(* IEC 61131-3 sources: 2026_Projet_YGO_ExcavatriceDragage/CODE/L_SIMULATION, 12 files *)

(* ---- FB_Sim_Encoder.st ---- *)
(* ═══════════════════════════════════════════════════════════════
   🧪 FB_Sim_Encoder — Simulation physique d'un codeur absolu de treuil
   ───────────────────────────────────────────────────────────────
   📄 Doc métier : DOC/AF/AF_Partie-13_Fonction_Simulation_v2.5.md
   📄 Spec composant : DOC/AF/AF_Partie-13_Fonction_Simulation/FB_Sim_Encoder_v1.1.md
   🧩 Brique réduite (Partie3 §1bis, "briques E/S & diagnostics") : pas de contrat
      Enable/Reset/Error complet, pas de StartStop/SafeStop — outil de banc, pas
      du métier machine.
   🎯 Rôle : fait "compter" un codeur absolu comme si le treuil tournait
      réellement, à partir des relais de sens commandés et du palier de vitesse courant.
   📥 Enable      : simulation active (SimulationModeActive AND NOT BusEncoderMxIsReal)
   📥 RelayFwd/RelayRev : sens commandé (contacteurs de sens du treuil)
   📥 StepNumber  : palier vitesse courant (1..5) — ex. instWinchM1.StepNumber
      Vitesse = interpolation linéaire : palier 1 → MinSpeedMps (1 m/s), palier 5 → MaxSpeedMps (2 m/s).
   📥 PresetCmd   : TRUE le cycle où un preset (homing) doit être appliqué (PresettTrigCmd = 2)
   📥 PresetValue : valeur brute à charger lors du preset
   📥 SpeedScaleFactor : facteur fin de confort (réglable à chaud, sans recompiler). Défaut 1.0 = vitesse
      réelle telle que définie par MinSpeedMps/MaxSpeedMps/PointsPerRev/CableM_PerRev/CycleTimeS.
   📤 RawPosOut   : position brute simulée (UDINT), à aiguiller à la place de la valeur
      EtherCAT réelle quand le device n'est pas Operational (voir PRG_02_Encoders.st)
   🔒 Comptage brut : entier SIGNÉ 32 bits (le conteneur UDINT n'est qu'un support d'échange,
      relu en DINT par toute la chaîne aval). Il franchit 0 sans jamais s'y figer ; la seule
      borne est la plage de représentation, signalée par CountSaturated — jamais muette.
   📤 CountSaturated : comptage en butée de plage du modèle (saturation signalée, vitesse purgée)
   `RawPos` en `VAR_IN_OUT`, référencé depuis `GVL_PERSISTENT`
      (même pattern que `Calib` dans `FB_Encoder_Homing`) — `PERSISTENT` n'est valide que sur du
      `VAR_GLOBAL` en CODESYS, pas sur une variable locale de FB. Un vrai codeur absolu physique
      conserve son comptage brut même à travers un reset FROID (indépendant de l'automate).
   ═══════════════════════════════════════════════════════════════ *)

// === DECLARATION (à coller dans la partie déclaration du POU FB_Sim_Encoder) ===

FUNCTION_BLOCK PUBLIC FB_Sim_Encoder
VAR_INPUT
    Enable           : BOOL;   (* --> [CMD] Active la simulation *)
    RelayFwd         : BOOL;   (* --> [HW] Sens commandé avant *)
    RelayRev         : BOOL;   (* --> [HW] Sens commandé arrière *)
    StepNumber       : INT;    (* --> [CMD] Palier vitesse courant (1..5, 0 = arrêt) *)
    PresetCmd        : BOOL;   (* --> [CMD] Applique un preset (homing) *)
    PresetValue      : UDINT;   (* --> [CFG] Valeur brute à charger au preset *)
    SpeedScaleFactor : REAL := 1.0;   (* --> [CFG] Facteur fin de confort (défaut 1.0) *)
    CoastDistanceM   : REAL := 0.0;   (* --> [CFG] Distance de roulis inertiel apres coupure des relais (m). 0 = arret net (defaut). >0 = le treuil continue a vitesse palier 1 dans le dernier sens sur CoastDistanceM metres -> modelise l'anticipation d'arret mecanique (ex. benne). *)
    PresetLatencyCycles : INT := 3;   (* --> [CFG] Nb cycles automate avant application du preset (referencement non instantane) *)
    TestOffsetCmd    : BOOL;          (* --> [TST] Front montant = applique TestOffsetPts (test banc) *)
    TestOffsetPts    : DINT := 0;     (* --> [TST] Décalage signé à appliquer (points bruts) *)
    // 📐 Paramètres physiques du treuil (mêmes valeurs que FB_Encoder_Scale) + vitesse réelle.
    // Vitesse simulée = interpolation linéaire du palier : palier 1 → MinSpeedMps, palier 5 → MaxSpeedMps.
    MinSpeedMps      : REAL := 1.0;    (* --> [CFG] Vitesse palier 1 (m/s) *)
    MaxSpeedMps      : REAL := 2.0;    (* --> [CFG] Vitesse palier 5 (m/s) *)
    PointsPerRev     : UDINT := 8192;  (* --> [CFG] Résolution codeur (pts/tour) *)
    CableM_PerRev    : REAL := 2.0;    (* --> [CFG] Développement câble (m/tour) *)
    CycleTimeS       : REAL := 0.010;  (* --> [CFG] Période tâche PLC (s) — MainTask 10 ms *)
    SpeedReportTauS  : REAL := 0.0;    (* --> [CFG][SYNTHETIQUE] Constante de temps 1er ordre du retour vitesse
        (RawSpdOut), s. 0.0 = saut instantane. >0 = RawSpdOut suit un 1er ordre vers la vitesse reelle du modele
        au lieu de sauter en escalier a la coupure des relais ; RawPosOut (position) n'est pas affecte. Valeur
        non calibree treuil M1/M2, plage indicative issue de la dynamique variateur M3 identifiee sur trace. *)
    // 🆕 Dynamique de glissement inertiel fidele (T421 cale sur trace reelle Suivi_86)
    CoastDecelUp_Mps2   : REAL := 1.20;  (* --> [CFG] Deceleration en montee (m/s²) : v0²/(2*0.543m) = 1.20 *)
    CoastDecelDown_Mps2 : REAL := 0.93;  (* --> [CFG] Deceleration en descente (m/s²) : v0²/(2*1.205m) = 0.93 *)
    MechanicStopEngaged : BOOL := FALSE; (* --> [HW] Butee mecanique engagee (coupe net le glissement) *)
END_VAR
VAR_OUTPUT
    RawPosOut   : UDINT;   (* <-- [DIAG] Position brute simulée *)
    RawSpdOut   : DINT;    (* <-- [DIAG] Vitesse brute simulée (0x6031:01 en 0.1 RPM) *)
    CountSaturated : BOOL; (* <-- [DIAG] Comptage en butée de plage du modèle (saturation signalée) *)
    CoastActive    : BOOL; (* <-- [DIAG] Indicateur de glissement inertiel en cours (T421) *)
END_VAR
VAR_IN_OUT
    RawPos      : UDINT;   (* <-> [BUS] Référence _SimEncoderRawPosM1/M2 (survit au reset froid) *)
END_VAR
VAR
    Increment        : UDINT;            (* . [LOC] Points ajoutés par cycle *)
    EffStep          : INT;              (* . [LOC] Pas borné (>= 1) *)
    SpeedMps         : REAL;             (* . [LOC] Vitesse simulée (m/s) *)
    TestOffsetEdge   : R_TRIG;           (* . [LOC] Front TestOffsetCmd *)
    PresetEdge       : R_TRIG;           (* . [LOC] Front montant PresetCmd *)
    PresetPending    : BOOL;             (* . [LOC] Preset en attente d'application (latence) *)
    PresetCount      : INT;              (* . [LOC] Compteur cycles de latence restants *)
    IncrStep1        : UDINT;            (* . [LOC] Increment par cycle a vitesse palier 1 (pour le roulis) *)
    MovingDir        : INT;              (* . [LOC] Dernier sens actif : +1 avant, -1 arriere, 0 arret *)
    CoastPtsLeft     : REAL;             (* . [LOC] Roulis inertiel restant (points bruts) *)
    TargetSpeedMps   : REAL;             (* . [LOC] Vitesse instantanee signee du modele position, avant filtrage retour *)
    ReportedSpeedMps : REAL;             (* . [LOC] Vitesse rapportee filtree 1er ordre, publiee dans RawSpdOut *)
    CoastSpeedMps    : REAL;             (* . [LOC] Vitesse instantanee signee pendant le glissement inertiel (T421) *)
END_VAR
VAR CONSTANT
    // 🛑 Plage de comptage du modèle : le compteur brut est un entier SIGNÉ 32 bits (le conteneur
    // UDINT n'est qu'un support d'échange, relu en DINT par toute la chaîne aval). La garde reste
    // volontairement à la moitié de la plage signée (2^30 pts = 262 144 m de câble) : inatteignable
    // en essai, elle interdit tout rebouclage silencieux si le modèle consommait toute sa plage.
    CST_CountTravelLimitPts : DINT := 1073741824; // 2^30 pts — demi-plage signée
END_VAR

// === IMPLEMENTATION (à coller dans le corps ST du POU FB_Sim_Encoder) ===

{region "§1 Gate"}
IF NOT Enable THEN
    RawPosOut := RawPos;
    // Comptage non evalue hors simulation : la saturation ne doit pas rester figee a TRUE.
    CountSaturated := FALSE;
    RETURN;
END_IF;
{endregion}

{region "§2 Injection test"}
// Injection test banc : VRAI saut de position (comme un glissement réel),
// pour tester Concept 1 / Méca E ET le rattrapage joystick (voir GVL_Simulation bandeau).
TestOffsetEdge(CLK := TestOffsetCmd);
IF TestOffsetEdge.Q THEN
    RawPos := DINT_TO_UDINT(UDINT_TO_DINT(RawPos) + TestOffsetPts);
END_IF;
{endregion}

{region "§3 Comptage"}
// 🎚️ Vitesse simulée = interpolation linéaire du palier (palier 1 → MinSpeedMps, palier 5 → MaxSpeedMps),
// pas par pas de (Max−Min)/4. Palier 0 (arrêt) ramène au palier 1 mais aucun mouvement n'est
// appliqué tant que RelayFwd/RelayRev = FALSE (section plus bas).
EffStep  := MAX(StepNumber, 1);
SpeedMps := MinSpeedMps + (INT_TO_REAL(EffStep) - 1.0) * ((MaxSpeedMps - MinSpeedMps) / 4.0);
// Points par cycle = vitesse (m/s) × points par mètre × période tâche (s) × facteur confort.
Increment := REAL_TO_UDINT(SpeedMps * (UDINT_TO_REAL(PointsPerRev) / CableM_PerRev) * CycleTimeS * SpeedScaleFactor);
// Increment "lent" (palier 1) : vitesse du roulis inertiel apres coupure des relais.
IncrStep1 := REAL_TO_UDINT(MinSpeedMps * (UDINT_TO_REAL(PointsPerRev) / CableM_PerRev) * CycleTimeS * SpeedScaleFactor);

// Front du preset : lance la latence de referencement (le codeur réel n'est pas
// instantane — il met PresetLatencyCycles cycles a se re-referencer apres le front).
PresetEdge(CLK := PresetCmd);
IF PresetEdge.Q THEN
    PresetPending := TRUE;
    PresetCount := PresetLatencyCycles;
END_IF;

// 📐 Le comptage brut est un entier SIGNÉ 32 bits : le conteneur UDINT n'est qu'un support
// d'échange (toute la chaîne aval le relit via UDINT_TO_DINT : FB_Encoder_Scale, FB_Encoder_Homing).
// Sa valeur 0 n'est donc PAS une butée mécanique — c'est un point de passage comme un autre, et
// c'est la seule façon de rester fidèle à un codeur absolu, dont le zéro de comptage est arbitraire.
// Aucune branche de comptage ne borne donc à un littéral : seule la garde de plage §3bis intervient,
// et elle est signalée (CountSaturated).
// Pendant l'attente du preset, la position brute est conservee (le codeur n'a pas encore re-reference).
// Le mouvement est gelé pendant la latence, comme un codeur réel en cours de referencement.
IF PresetPending THEN
    IF PresetCount > 0 THEN
        PresetCount := PresetCount - 1;
    ELSE
        // Latence écoulée : applique la valeur cible du preset.
        RawPos := PresetValue;
        PresetPending := FALSE;
    END_IF;
    TargetSpeedMps := 0.0;
ELSIF RelayFwd AND NOT RelayRev THEN
    IF NOT MechanicStopEngaged THEN
        RawPos := DINT_TO_UDINT(UDINT_TO_DINT(RawPos) + UDINT_TO_DINT(Increment));
        MovingDir := 1;
        CoastSpeedMps := SpeedMps;
        CoastPtsLeft := CoastDistanceM * (UDINT_TO_REAL(PointsPerRev) / CableM_PerRev);
        TargetSpeedMps := SpeedMps;
    ELSE
        MovingDir := 0;
        CoastSpeedMps := 0.0;
        CoastPtsLeft := 0.0;
        TargetSpeedMps := 0.0;
    END_IF;
    CoastActive := FALSE;
ELSIF RelayRev AND NOT RelayFwd THEN
    IF NOT MechanicStopEngaged THEN
        RawPos := DINT_TO_UDINT(UDINT_TO_DINT(RawPos) - UDINT_TO_DINT(Increment));
        MovingDir := -1;
        CoastSpeedMps := -SpeedMps;
        CoastPtsLeft := CoastDistanceM * (UDINT_TO_REAL(PointsPerRev) / CableM_PerRev);
        TargetSpeedMps := -SpeedMps;
    ELSE
        MovingDir := 0;
        CoastSpeedMps := 0.0;
        CoastPtsLeft := 0.0;
        TargetSpeedMps := 0.0;
    END_IF;
    CoastActive := FALSE;
ELSE
    // Relais coupes (ou les deux actifs = conflit) : glissement inertiel (T421)
    IF MechanicStopEngaged THEN
        MovingDir := 0;
        CoastSpeedMps := 0.0;
        CoastPtsLeft := 0.0;
        TargetSpeedMps := 0.0;
        CoastActive := FALSE;
    ELSIF (CoastDistanceM > 0.0) AND (CoastPtsLeft >= 1.0) AND (MovingDir <> 0) THEN
        // Mode historique compatibilite (si CoastDistanceM explicitement configure > 0)
        CoastActive := TRUE;
        IF MovingDir = 1 THEN
            RawPos := DINT_TO_UDINT(UDINT_TO_DINT(RawPos) + UDINT_TO_DINT(IncrStep1));
            TargetSpeedMps := MinSpeedMps;
        ELSE
            RawPos := DINT_TO_UDINT(UDINT_TO_DINT(RawPos) - UDINT_TO_DINT(IncrStep1));
            TargetSpeedMps := -MinSpeedMps;
        END_IF;
        CoastPtsLeft := CoastPtsLeft - UDINT_TO_REAL(IncrStep1);
    ELSIF (ABS(CoastSpeedMps) > 0.005) AND (MovingDir <> 0) THEN
        // 🆕 Modele dynamique continu T421 : deceleration signee continue calee sur trace reelle
        CoastActive := TRUE;
        IF CoastSpeedMps > 0.0 THEN
            CoastSpeedMps := CoastSpeedMps - CoastDecelUp_Mps2 * CycleTimeS;
            IF CoastSpeedMps <= 0.005 THEN
                CoastSpeedMps := 0.0;
                MovingDir := 0;
                CoastActive := FALSE;
            END_IF;
        ELSE
            CoastSpeedMps := CoastSpeedMps + CoastDecelDown_Mps2 * CycleTimeS;
            IF CoastSpeedMps >= -0.005 THEN
                CoastSpeedMps := 0.0;
                MovingDir := 0;
                CoastActive := FALSE;
            END_IF;
        END_IF;

        // Deplacement par cycle correspondant a CoastSpeedMps
        Increment := REAL_TO_UDINT(ABS(CoastSpeedMps) * (UDINT_TO_REAL(PointsPerRev) / CableM_PerRev) * CycleTimeS * SpeedScaleFactor);
        IF CoastSpeedMps > 0.0 THEN
            RawPos := DINT_TO_UDINT(UDINT_TO_DINT(RawPos) + UDINT_TO_DINT(Increment));
            TargetSpeedMps := CoastSpeedMps;
        ELSIF CoastSpeedMps < 0.0 THEN
            RawPos := DINT_TO_UDINT(UDINT_TO_DINT(RawPos) - UDINT_TO_DINT(Increment));
            TargetSpeedMps := CoastSpeedMps;
        ELSE
            TargetSpeedMps := 0.0;
        END_IF;
    ELSE
        MovingDir := 0;
        CoastSpeedMps := 0.0;
        CoastPtsLeft := 0.0;
        TargetSpeedMps := 0.0;
        CoastActive := FALSE;
    END_IF;
END_IF;
{endregion}

{region "§3bis Garde de plage de comptage"}
// 🛑 SEULE borne du comptage : la plage de représentation signée. Elle est SIGNALÉE
// (CountSaturated) et cohérente — une position bornée ne publie plus de vitesse de mouvement,
// ce qui interdit la signature « position figée + vitesse non nulle + zéro défaut ».
CountSaturated := FALSE;
IF UDINT_TO_DINT(RawPos) > CST_CountTravelLimitPts THEN
    RawPos := DINT_TO_UDINT(CST_CountTravelLimitPts);
    CountSaturated := TRUE;
ELSIF UDINT_TO_DINT(RawPos) < -CST_CountTravelLimitPts THEN
    RawPos := DINT_TO_UDINT(-CST_CountTravelLimitPts);
    CountSaturated := TRUE;
END_IF;
IF CountSaturated THEN
    TargetSpeedMps := 0.0;
END_IF;
{endregion}

{region "§4 Sortie"}
RawPosOut := RawPos;
// Retour vitesse rapporte (RawSpdOut) : 1er ordre vers TargetSpeedMps. SpeedReportTauS=0.0
// -> alpha=1 -> saut instantane (comportement historique inchange).
ReportedSpeedMps := ReportedSpeedMps
    + (CycleTimeS / (SpeedReportTauS + CycleTimeS)) * (TargetSpeedMps - ReportedSpeedMps);
// Formule inverse vitesse brute EtherCAT CoE (0.1 RPM) :
// SpdValue = (V_mps * 60.0) / (0.1 * CableM_PerRev) = V_mps * 300.0 (sur tambour 2m)
IF (CableM_PerRev > 0.0) THEN
    RawSpdOut := REAL_TO_DINT((ReportedSpeedMps * 60.0) / (0.1 * CableM_PerRev) * SpeedScaleFactor);
ELSE
    RawSpdOut := 0;
END_IF;
{endregion}

END_FUNCTION_BLOCK

(* ---- FB_Sim_Joystick.st ---- *)
(* =======================================================================
   🧪 FB_Sim_Joystick — Simulation des entrees brutes joystick (bus CAN hors ligne)
   🎯 Rôle : reproduire un geste operateur depuis un bouton directionnel.
   Appui armement, debattement, relachement armement, retour dynamique.
   Aucun etat arme produit ; permis et armement restent au joystick reel.
   📄 Doc métier : DOC/AF/AF_Partie-13_Fonction_Simulation_v2.5.md
   ======================================================================= *)

// === DECLARATION (à coller dans la partie déclaration du POU FB_Sim_Joystick) ===

FUNCTION_BLOCK PUBLIC FB_Sim_Joystick
VAR_INPUT
    Enable              : BOOL;   (* --> [CMD] Active la simulation *)
    NeutralRaw          : INT := 5000;   (* --> [CFG] Valeur brute au repos (neutre) *)
    MaxRaw              : INT := 10000;   (* --> [CFG] Valeur brute à fond *)
    BtnLeft_Rev_TREMIE  : BOOL;   (* --> [TST] Bouton gauche : X→0, Y→neutre *)
    BtnRight_Fwd_MAINT  : BOOL;   (* --> [TST] Bouton droite : X→MaxRaw, Y→neutre *)
    BtnFwd_Up_Close     : BOOL;   (* --> [TST] Bouton avant : X→neutre, Y→MaxRaw *)
    BtnRev_Down_Open    : BOOL;   (* --> [TST] Bouton arrière : X→neutre, Y→0 *)
    OvershootActive     : BOOL;   (* --> [TST] Dépassement de montée au-delà de 100% (défaut capteur hors plage) *)
    BagotementActive    : BOOL;   (* --> [TST] Bagotement au relâchement (petit balancement autour du neutre) *)
    RiseTimeS           : REAL := 1.5;   (* --> [CFG] Temps de montée 0→100% (s) *)
    FallTimeMs          : TIME := T#200MS;   (* --> [CFG] Temps de retombée 100%→0 *)
    CycleTimeS          : REAL := 0.010;   (* --> [CFG] Période tâche PLC (s) — 10 ms *)
    GesturePermit       : BOOL := TRUE; (* --> [SAFE] Stimuli manuels au repos avant un geste automatique *)
    ArmHoldTime         : TIME := T#200MS; (* --> [CFG] Appui bouton avant debattement *)
    ButtonReleaseDelay  : TIME := T#200MS; (* --> [CFG] Maintien bouton apres debut debattement *)
END_VAR
VAR_OUTPUT
    RawX        : INT;   (* <-- [DIAG] Valeur brute axe X (dynamique, neutre = NeutralRaw) *)
    RawY        : INT;   (* <-- [DIAG] Valeur brute axe Y (dynamique, neutre = NeutralRaw) *)
    RawButton   : BOOL;  (* <-- [DIAG] Appui armement simule, relache pendant le maintien du manche *)
    ModelActive : BOOL;  (* <-- [STAT] Propriete exclusive des trois entrees brutes pendant le geste et le retour *)
    ReturningActive : BOOL;  (* <-- [STAT] TRUE si retour dynamique en cours (FALL/OVERSHOOT) — FB_SimBench émet le modèle *)
END_VAR
VAR
    instArmTimer : TON; (* * [INST] Maintien armement avant debattement *)
    instButtonReleaseTimer : TON; (* * [INST] Relachement bouton apres debut debattement *)
    GestureStep : INT := 0; (* . [LOC] Attente relachement, disponible, appui, mouvement *)
    RequestedDirection : INT; (* . [LOC] Direction unique demandee, 0 si aucune ou conflit *)
    GestureDirection : INT; (* . [LOC] Direction memorisee au nouvel appui *)
    DeflectionActive : BOOL; (* . [LOC] Debattement admis pour le geste courant *)
    RequestMatchesGesture : BOOL; (* . [LOC] Direction demandee identique au geste *)
    TimingValid : BOOL; (* . [LOC] Parametres dynamiques strictement positifs *)
    FirstCycle  : BOOL := TRUE;   (* . [LOC] Initialisation au neutre *)
    State       : INT := 0;   (* . [LOC] 0=IDLE, 1=RISE, 2=FALL, 3=OVERSHOOT *)
    TargetX     : INT;   (* . [LOC] Cible brute axe X *)
    TargetY     : INT;   (* . [LOC] Cible brute axe Y *)
    ActiveAxis  : INT;   (* . [LOC] 0=aucun, 1=X, 2=Y (axe en retour) *)
    RiseStep    : REAL;   (* . [LOC] Pas de montée par cycle (points) *)
    FallStep    : REAL;   (* . [LOC] Pas de retombée par cycle (points) *)
    RandCnt     : INT := 0;   (* . [LOC] Compteur pseudo-aléatoire (bruit de montée) *)
    Noise       : INT;   (* . [LOC] Bruit ±25 points (≈ ±0.5% de la course) *)
    BtnCount    : INT;   (* . [LOC] Nombre de boutons directionnels actifs (0..4) *)
    OscDev      : REAL;   (* . [LOC] Écart au neutre de l'oscillateur de bagotement *)
    OscVel      : REAL;   (* . [LOC] Vitesse de l'oscillateur (points/cycle) *)
    OscAcc      : REAL;   (* . [LOC] Accélération de l'oscillateur *)
END_VAR
VAR CONSTANT
    CST_GESTURE_WAIT_RELEASE : INT := 0; (* . [CFG] Relachement complet et retour neutre requis *)
    CST_GESTURE_READY : INT := 1; (* . [CFG] Nouveau geste disponible *)
    CST_GESTURE_ARM : INT := 2; (* . [CFG] Appui armement, manche neutre *)
    CST_GESTURE_MOVE : INT := 3; (* . [CFG] Manche deplace, bouton ensuite relache *)
    CST_DIRECTION_LEFT : INT := 1; (* . [CFG] Demande X negatif *)
    CST_DIRECTION_RIGHT : INT := 2; (* . [CFG] Demande X positif *)
    CST_DIRECTION_FORWARD : INT := 3; (* . [CFG] Demande Y positif *)
    CST_DIRECTION_REVERSE : INT := 4; (* . [CFG] Demande Y negatif *)
    CST_ST_IDLE      : INT := 0;   (* . [CFG] État : au neutre *)
    CST_ST_RISE      : INT := 1;   (* . [CFG] État : montée vers la cible *)
    CST_ST_FALL      : INT := 2;   (* . [CFG] État : retombée linéaire *)
    CST_ST_OVERSHOOT : INT := 3;   (* . [CFG] État : bagotement (oscillations amorties) *)
    CST_OSC_K        : REAL := 0.01;   (* . [CFG] Raideur oscillateur (fréquence bagotement) *)
    CST_OSC_C        : REAL := 0.05;   (* . [CFG] Amortissement (2-3 oscillations visibles) *)
    CST_OVERSHOOT_AMT : INT := 600;   (* . [CFG] Dépassement de montée au-delà de MaxRaw (déclenche défaut capteur hors plage) *)
    CST_BAGOT_AMT     : INT := 500;   (* . [CFG] Amplitude du bagotement au relâchement (~5% autour du neutre) *)
END_VAR

// === IMPLEMENTATION (à coller dans le corps ST du POU FB_Sim_Joystick) ===

{region "§1 Gate"}
// 🔑 Initialise au neutre au premier cycle uniquement ; ensuite RawX/RawY sont pilotés
// dynamiquement par les boutons. Quand la simulation est coupée, on revient au neutre.
TimingValid := (RiseTimeS > 0.0) AND (CycleTimeS > 0.0) AND (FallTimeMs > T#0MS);
IF NOT Enable OR NOT TimingValid THEN
    FirstCycle := TRUE;
    State      := CST_ST_IDLE;
    RawX       := NeutralRaw;
    RawY       := NeutralRaw;
    RawButton  := FALSE;
    ReturningActive := FALSE; // 📊 Neutralisation : simulation inactive hors Enable
    ModelActive := FALSE;
    GestureStep := CST_GESTURE_WAIT_RELEASE;
    GestureDirection := 0;
    instArmTimer(IN := FALSE, PT := ArmHoldTime);
    instButtonReleaseTimer(IN := FALSE, PT := ButtonReleaseDelay);
    RETURN;
END_IF;
{endregion}

{region "§2 Initialisation neutre"}
IF FirstCycle THEN
    RawX       := NeutralRaw;
    RawY       := NeutralRaw;
    RawButton  := FALSE;
    State      := CST_ST_IDLE;
    FirstCycle := FALSE;
    GestureStep := CST_GESTURE_WAIT_RELEASE;
END_IF;
{endregion}

{region "§3 Pseudo-aléatoire (bruit de montée)"}
// 🎲 Compteur qui repasse à zéro, multiplié pour rester dans la plage (méthode validée).
// Le bruit s'ajoute à la rampe de montée uniquement (pas à la retombée, linéaire propre).
RandCnt := (RandCnt + 1) MOD 1000;
Noise   := (RandCnt MOD 50) - 25;   // ±25 points (≈ ±0.5% de la course)
{endregion}

{region "§4 Cibles & transitions"}
// 🎯 Un SEUL bouton impose une butée d'axe ; 0 ou ≥2 boutons = neutre (pas de diagonale implicite).
// Si OvershootActive : la cible de montée DÉPASSE la butée (MaxRaw+AMT ou 0−AMT) pour
// déclencher le défaut capteur hors plage (RawOutOfRange) — test du dépassement de valeur.
BtnCount := BOOL_TO_INT(BtnLeft_Rev_TREMIE) + BOOL_TO_INT(BtnRight_Fwd_MAINT)
          + BOOL_TO_INT(BtnFwd_Up_Close) + BOOL_TO_INT(BtnRev_Down_Open);
RequestedDirection := 0;
IF BtnCount = 1 THEN
    IF BtnLeft_Rev_TREMIE THEN RequestedDirection := CST_DIRECTION_LEFT;
    ELSIF BtnRight_Fwd_MAINT THEN RequestedDirection := CST_DIRECTION_RIGHT;
    ELSIF BtnFwd_Up_Close THEN RequestedDirection := CST_DIRECTION_FORWARD;
    ELSE RequestedDirection := CST_DIRECTION_REVERSE;
    END_IF;
END_IF;

// Un seul appui brut par geste ; aucun nouvel essai tant que l'IHM reste tenue.
instArmTimer(IN := GestureStep = CST_GESTURE_ARM, PT := ArmHoldTime);
instButtonReleaseTimer(IN := GestureStep = CST_GESTURE_MOVE, PT := ButtonReleaseDelay);
DeflectionActive := FALSE;
RawButton := FALSE;
RequestMatchesGesture := (RequestedDirection = GestureDirection) AND (BtnCount = 1);
IF BtnCount > 0 THEN ModelActive := TRUE; END_IF;
IF NOT GesturePermit THEN GestureStep := CST_GESTURE_WAIT_RELEASE; END_IF;

IF GestureStep = CST_GESTURE_WAIT_RELEASE THEN
        // Les boutons doivent etre relaches APRES stabilisation du retour.
        IF (BtnCount = 0) AND (State = CST_ST_IDLE) AND GesturePermit THEN
            GestureStep := CST_GESTURE_READY;
            ModelActive := FALSE;
        END_IF;
ELSIF GestureStep = CST_GESTURE_READY THEN
        IF BtnCount = 1 THEN
            GestureDirection := RequestedDirection;
            GestureStep := CST_GESTURE_ARM;
            RawButton := TRUE;
        ELSIF BtnCount > 1 THEN
            GestureStep := CST_GESTURE_WAIT_RELEASE;
        END_IF;
ELSIF GestureStep = CST_GESTURE_ARM THEN
        IF NOT RequestMatchesGesture THEN
            GestureStep := CST_GESTURE_WAIT_RELEASE;
        ELSE
            RawButton := TRUE;
            IF instArmTimer.Q THEN GestureStep := CST_GESTURE_MOVE; END_IF;
        END_IF;
ELSIF GestureStep = CST_GESTURE_MOVE THEN
        IF NOT RequestMatchesGesture THEN
            GestureStep := CST_GESTURE_WAIT_RELEASE;
        ELSE
            DeflectionActive := TRUE;
            RawButton := NOT instButtonReleaseTimer.Q;
        END_IF;
ELSE
    GestureStep := CST_GESTURE_WAIT_RELEASE;
END_IF;

IF DeflectionActive THEN
    IF BtnLeft_Rev_TREMIE THEN
        IF OvershootActive THEN TargetX := 0 - CST_OVERSHOOT_AMT; ELSE TargetX := 0; END_IF;
        TargetY := NeutralRaw; ActiveAxis := 1;
    ELSIF BtnRight_Fwd_MAINT THEN
        IF OvershootActive THEN TargetX := MaxRaw + CST_OVERSHOOT_AMT; ELSE TargetX := MaxRaw; END_IF;
        TargetY := NeutralRaw; ActiveAxis := 1;
    ELSIF BtnFwd_Up_Close THEN
        TargetX := NeutralRaw;
        IF OvershootActive THEN TargetY := MaxRaw + CST_OVERSHOOT_AMT; ELSE TargetY := MaxRaw; END_IF;
        ActiveAxis := 2;
    ELSE
        TargetX := NeutralRaw;
        IF OvershootActive THEN TargetY := 0 - CST_OVERSHOOT_AMT; ELSE TargetY := 0; END_IF;
        ActiveAxis := 2;
    END_IF;
    State := CST_ST_RISE;
ELSE
    // 0 ou ≥2 boutons : retour au neutre.
    TargetX := NeutralRaw;
    TargetY := NeutralRaw;
    IF State = CST_ST_RISE THEN
        // Front de relâchement : retour au neutre. D'abord retombée linéaire (FALL),
        // puis petit bagotement de quelques % autour du neutre si OvershootActive (voir §6).
        State := CST_ST_FALL;
    END_IF;
END_IF;
{endregion}

{region "§5 Ascending (rampe + bruit)"}
IF State = CST_ST_RISE THEN
    // Pas de montée : pleine course (MaxRaw−NeutralRaw) en RiseTimeS.
    RiseStep := INT_TO_REAL(MaxRaw - NeutralRaw) / (RiseTimeS / CycleTimeS);
    // Axe X
    IF RawX < TargetX THEN
        RawX := MIN(RawX + REAL_TO_INT(RiseStep) + Noise, TargetX);
    ELSIF RawX > TargetX THEN
        RawX := MAX(RawX - REAL_TO_INT(RiseStep) - Noise, TargetX);
    END_IF;
    // Axe Y
    IF RawY < TargetY THEN
        RawY := MIN(RawY + REAL_TO_INT(RiseStep) + Noise, TargetY);
    ELSIF RawY > TargetY THEN
        RawY := MAX(RawY - REAL_TO_INT(RiseStep) - Noise, TargetY);
    END_IF;
END_IF;
{endregion}

{region "§6 Retombée linéaire (sans bagotement)"}
IF State = CST_ST_FALL THEN
    // Pas de retombée : pleine course en FallTimeMs (TIME_TO_REAL → ms, /1000 → s).
    FallStep := INT_TO_REAL(MaxRaw - NeutralRaw) / (TIME_TO_REAL(FallTimeMs) / 1000.0 / CycleTimeS);
    IF RawX < NeutralRaw THEN
        RawX := MIN(RawX + REAL_TO_INT(FallStep), NeutralRaw);
    ELSIF RawX > NeutralRaw THEN
        RawX := MAX(RawX - REAL_TO_INT(FallStep), NeutralRaw);
    END_IF;
    IF RawY < NeutralRaw THEN
        RawY := MIN(RawY + REAL_TO_INT(FallStep), NeutralRaw);
    ELSIF RawY > NeutralRaw THEN
        RawY := MAX(RawY - REAL_TO_INT(FallStep), NeutralRaw);
    END_IF;
    IF RawX = NeutralRaw AND RawY = NeutralRaw THEN
        // Arrivée au neutre : si bagotement demandé, lance un petit balancement de quelques %.
        IF BagotementActive THEN
            State := CST_ST_OVERSHOOT;
            IF ActiveAxis = 1 THEN
                OscDev := INT_TO_REAL(CST_BAGOT_AMT);
            ELSE
                OscDev := INT_TO_REAL(CST_BAGOT_AMT);
            END_IF;
            OscVel := 0.0;
        ELSE
            State := CST_ST_IDLE;
        END_IF;
    END_IF;
END_IF;
{endregion}

{region "§7 Bagotement (dépassement + oscillations amorties)"}
IF State = CST_ST_OVERSHOOT THEN
    // 🎢 Oscillateur harmonique amorti discret (semi-implicite) autour du neutre :
    // le joystick dépasse le centre (~12% de l'écart initial) puis oscille 1-2 fois
    // avant de se stabiliser — comportement d'un opérateur qui relâche et balance.
    OscAcc := -CST_OSC_K * OscDev - CST_OSC_C * OscVel;
    OscVel := OscVel + OscAcc;
    OscDev := OscDev + OscVel;
    IF ActiveAxis = 1 THEN
        RawX := NeutralRaw + REAL_TO_INT(OscDev);
    ELSE
        RawY := NeutralRaw + REAL_TO_INT(OscDev);
    END_IF;
    // Stabilisé : revient exactement au centre.
    IF ABS(OscDev) < 1.0 AND ABS(OscVel) < 1.0 THEN
        State := CST_ST_IDLE;
        IF ActiveAxis = 1 THEN
            RawX := NeutralRaw;
        ELSE
            RawY := NeutralRaw;
        END_IF;
    END_IF;
END_IF;
{endregion}

{region "§8 Homme-mort brut + drapeau retour"}
// RawButton est exclusivement produit par le sequenceur du geste (§4).
// Drapeau "retour dynamique en cours" : TRUE si l'état est FALL ou OVERSHOOT (retombée/bagotement).
// Permet à FB_SimBench d'émettre la sortie du modèle même après relâchement du bouton.
ReturningActive := (State = CST_ST_FALL) OR (State = CST_ST_OVERSHOOT);
{endregion}

END_FUNCTION_BLOCK

(* ---- FB_Sim_KlossTorque.st ---- *)
(* ═══════════════════════════════════════════════════════════════
   🧪 FB_Sim_KlossTorque — Couple electromagnetique, formule de Kloss
   ───────────────────────────────────────────────────────────────
   🎯 Role : Calcul factorise du couple moteur asynchrone (Kloss), reutilise
   par le regime etabli et le test de decrochage a glissement bloque.
   📄 Doc metier : DOC/WFLOW/CONTRACTS/PLAN_T317_SIMBENCH_TREUIL_ELECTRIQUE.md
   🧩 Dependances : aucune (calcul pur)
   ═══════════════════════════════════════════════════════════════ *)
FUNCTION_BLOCK PUBLIC FB_Sim_KlossTorque
VAR_INPUT
    // === CONTRAT LIGHT ===
    Enable                 : BOOL; // --> [CMD] Autorisation generale FB

    // === CALCUL ===
    MaxTorque_Nm           : REAL; // --> [CFG] Cmax decrochage
    Slip_Ratio              : REAL; // --> [CMD] Glissement (jamais 0.0 -- protege par l'appelant)
    SlipAtMaxTorque_Ratio   : REAL; // --> [CFG] gmax au point de fonctionnement courant
    VoltageRatio2           : REAL := 1.0; // --> [CMD] (U_act/U_nom)^2
END_VAR
VAR_OUTPUT
    Ready                  : BOOL; // <-- [STAT] FB pret
    Torque_Nm              : REAL; // <-- [DIAG] Couple electromagnetique resultant
END_VAR

IF NOT Enable THEN
    Ready := FALSE;
    Torque_Nm := 0.0;
    RETURN;
END_IF;

Torque_Nm := 2.0 * MaxTorque_Nm
    / (Slip_Ratio / SlipAtMaxTorque_Ratio + SlipAtMaxTorque_Ratio / Slip_Ratio)
    * VoltageRatio2;

Ready := TRUE;

(* ---- FB_Sim_PositionSensor.st ---- *)
(* DOC: DOC/AF/AF_Partie-13_Fonction_Simulation_v2.5.md
   Capteur de position cumulatif avec hysteresis et episode intermittent rejouable.
   Cette brique ne connait ni le mouvement ni la logique M3 : elle transforme uniquement
   une position mecanique vraie en DI. *)
FUNCTION_BLOCK PUBLIC FB_Sim_PositionSensor
VAR_INPUT
    Enable : BOOL;
    Position_M : REAL;
    Threshold_M : REAL;
    Hysteresis_M : REAL := 0.02;
    ActiveBelowThreshold : BOOL := TRUE;
    ElectricalDelayS : REAL := 0.0;
    IntermittenceActive : BOOL := FALSE;
    IntermittenceDurationS : REAL := 1.0;
    IntermittencePeriodS : REAL := 0.12;
    ScenarioSeed : UDINT := 1;
    CycleTimeS : REAL := 0.01;
    (* Profil « BLIP COURT » — SECOND profil, independant du train de bascules du profil
       d'intermittence ci-dessus (dont les parametres restent inchanges).
       0 = desactive : le comportement historique est strictement conserve.
       Rejoue les excursions electriques courtes mesurees sur la trace terrain du
       2026-09-04 : Tremie contradictoire pendant 2 echantillons a 12,24 s (~200 ms) et
       PV reactive 1 echantillon a 14,94 s (~100 ms).
         BlipTransitions = nombre de bascules electriques (1 = une excursion puis retour) ;
         BlipDurationS   = duree de maintien de chaque etat, donc largeur de l'excursion. *)
    BlipTransitions : UDINT := 0;
    BlipDurationS : REAL := 0.2;
    (* L5 (2026-10-28) — MECANISME DE CAME, SPATIAL : en franchissant le capteur on le VOIT,
       on le PERD sur une courte zone, on le RETROUVE, puis il reste FIXE. Lie a la POSITION
       (pas au temps) : se produit a chaque passage, dans les DEUX sens, et reste stable a
       l'arret (bornes de la zone avec hysteresis CST_CamHysteresis_M contre le bruit/balancement).
       Zone de perte placee APRES le front de detection (cote -/+ Hysteresis_M) :
       [front - Start - Width ; front - Start] cote detection.
       FALSE = historique strictement inchange. Valeurs = HYPOTHESES. *)
    CamDropoutActive : BOOL := FALSE;
    CamDropoutStart_M : REAL := 0.02;
    CamDropoutWidth_M : REAL := 0.04;
    (* Came finie : FALSE = capteur cumulatif ; TRUE = sortie active uniquement sur CamLength_M apres Threshold_M. *)
    FiniteCamActive : BOOL := FALSE;
    CamLength_M : REAL := 0.0;
END_VAR
VAR_OUTPUT
    RawDetected : BOOL;
    ElectricalOutput : BOOL;
    EpisodeActive : BOOL;
    BlipActive : BOOL;
    TransitionCount : UDINT;
    EpisodeTogglePeriodS : REAL;
END_VAR
VAR
    Initialized : BOOL;
    PreviousRawDetected : BOOL;
    EpisodeTarget : BOOL;
    DelayTimerS : REAL;
    EpisodeTimerS : REAL;
    ToggleTimerS : REAL;
    RandomState : UDINT;
    BlipRunning : BOOL;
    BlipTimerS : REAL;
    BlipCount : UDINT;
    HystDetected : BOOL;      (* L5 : etat mecanique avec hysteresis (avant perte de came) *)
    InCamDropout : BOOL;      (* L5 : position dans la zone de perte de la came *)
    CamNear_M : REAL;         (* L5 : borne de la zone cote front de detection *)
    CamFar_M : REAL;          (* L5 : borne de la zone cote interieur *)
    PastFiniteCam : BOOL;     (* Depassement au-dela de la longueur physique de came *)
    CamEnd_M : REAL;          (* Borne de fin de came finie *)
END_VAR
VAR CONSTANT
    (* Plafond du nombre de bascules du profil « blip court » : borne la duree de l'episode
       et interdit tout rebouclage de compteur UDINT (revue du 2026-09-20, F9). *)
    CST_BlipMaxTransitions : UDINT := 1000;
    CST_CamHysteresis_M : REAL := 0.01;   (* L5 : hysteresis des bornes de la zone de perte *)
END_VAR

IF NOT Enable THEN
    Initialized := FALSE;
    RawDetected := FALSE;
    ElectricalOutput := FALSE;
    PreviousRawDetected := FALSE;
    EpisodeActive := FALSE;
    BlipActive := FALSE;
    BlipRunning := FALSE;
    BlipTimerS := 0.0;
    BlipCount := 0;
    DelayTimerS := 0.0;
    EpisodeTimerS := 0.0;
    ToggleTimerS := 0.0;
    TransitionCount := 0;
    EpisodeTogglePeriodS := 0.0;
    PastFiniteCam := FALSE;
    RETURN;
END_IF;

(* Hysteresis sur une frontiere cumulative : les cinq DI restent compatibles avec
   le mot thermometre du decodeur M3, contrairement a cinq fenetres independantes. *)
IF NOT Initialized THEN
    IF ActiveBelowThreshold THEN
        RawDetected := Position_M <= Threshold_M;
        IF FiniteCamActive THEN
            PastFiniteCam := Position_M < (Threshold_M - MAX(0.0, CamLength_M));
            RawDetected := RawDetected AND NOT PastFiniteCam;
        ELSE
            PastFiniteCam := FALSE;
        END_IF;
    ELSE
        RawDetected := Position_M >= Threshold_M;
        IF FiniteCamActive THEN
            PastFiniteCam := Position_M > (Threshold_M + MAX(0.0, CamLength_M));
            RawDetected := RawDetected AND NOT PastFiniteCam;
        ELSE
            PastFiniteCam := FALSE;
        END_IF;
    END_IF;
    HystDetected := RawDetected;
    ElectricalOutput := RawDetected;
    PreviousRawDetected := RawDetected;
    RandomState := ScenarioSeed MOD 1000000;
    IF RandomState = 0 THEN
        RandomState := 1;
    END_IF;
    EpisodeTogglePeriodS := MAX(0.01, IntermittencePeriodS);
    Initialized := TRUE;
    RETURN;
END_IF;

IF ActiveBelowThreshold THEN
    IF HystDetected THEN
        HystDetected := Position_M <= (Threshold_M + MAX(0.0, Hysteresis_M));
    ELSE
        HystDetected := Position_M <= (Threshold_M - MAX(0.0, Hysteresis_M));
    END_IF;
    (* Zone de perte : apres le front d'entree en detection (cote - hysteresis), vers l'interieur. *)
    CamNear_M := Threshold_M - MAX(0.0, Hysteresis_M) - MAX(0.0, CamDropoutStart_M);
    CamFar_M := CamNear_M - MAX(0.0, CamDropoutWidth_M);
    IF NOT CamDropoutActive THEN
        InCamDropout := FALSE;
    ELSIF InCamDropout THEN
        InCamDropout := (Position_M <= CamNear_M + CST_CamHysteresis_M) AND (Position_M > CamFar_M - CST_CamHysteresis_M);
    ELSE
        InCamDropout := (Position_M <= CamNear_M - CST_CamHysteresis_M) AND (Position_M > CamFar_M + CST_CamHysteresis_M);
    END_IF;
    CamEnd_M := Threshold_M - MAX(0.0, CamLength_M);
    IF NOT FiniteCamActive THEN
        PastFiniteCam := FALSE;
    ELSIF PastFiniteCam THEN
        PastFiniteCam := Position_M < (CamEnd_M + CST_CamHysteresis_M);
    ELSE
        PastFiniteCam := Position_M < CamEnd_M;
    END_IF;
ELSE
    IF HystDetected THEN
        HystDetected := Position_M >= (Threshold_M - MAX(0.0, Hysteresis_M));
    ELSE
        HystDetected := Position_M >= (Threshold_M + MAX(0.0, Hysteresis_M));
    END_IF;
    CamNear_M := Threshold_M + MAX(0.0, Hysteresis_M) + MAX(0.0, CamDropoutStart_M);
    CamFar_M := CamNear_M + MAX(0.0, CamDropoutWidth_M);
    IF NOT CamDropoutActive THEN
        InCamDropout := FALSE;
    ELSIF InCamDropout THEN
        InCamDropout := (Position_M >= CamNear_M - CST_CamHysteresis_M) AND (Position_M < CamFar_M + CST_CamHysteresis_M);
    ELSE
        InCamDropout := (Position_M >= CamNear_M + CST_CamHysteresis_M) AND (Position_M < CamFar_M - CST_CamHysteresis_M);
    END_IF;
    CamEnd_M := Threshold_M + MAX(0.0, CamLength_M);
    IF NOT FiniteCamActive THEN
        PastFiniteCam := FALSE;
    ELSIF PastFiniteCam THEN
        PastFiniteCam := Position_M > (CamEnd_M - CST_CamHysteresis_M);
    ELSE
        PastFiniteCam := Position_M > CamEnd_M;
    END_IF;
END_IF;
(* L5 : perte de came + came finie ; hors options, RawDetected = HystDetected. *)
RawDetected := HystDetected AND NOT InCamDropout AND NOT PastFiniteCam;

(* Un episode est declenche par un franchissement mecanique, pas par une de ses
   propres bascules electriques. Les fronts restent donc bornes et reproductibles. *)
IF RawDetected <> PreviousRawDetected THEN
    PreviousRawDetected := RawDetected;
    EpisodeTarget := RawDetected;
    (* Une bascule mecanique pendant l'episode modifie seulement la cible finale.
       Elle ne remet jamais son chronometre a zero : l'episode reste borne. *)
    IF NOT EpisodeActive THEN
        DelayTimerS := 0.0;
        EpisodeTimerS := 0.0;
        ToggleTimerS := 0.0;
        (* Tirage unique par episode : reproductible pour une graine et sans bruit
           blanc scan-par-scan. La periode varie de 70 % a 130 % du nominal. *)
        RandomState := RandomState + 7919;
        IF RandomState >= 1000000 THEN
            RandomState := RandomState - 1000000;
        END_IF;
        EpisodeTogglePeriodS := MAX(0.01, IntermittencePeriodS
            * (0.7 + UDINT_TO_REAL(RandomState MOD 6000) / 10000.0));
        EpisodeActive := IntermittenceActive AND (IntermittenceDurationS > 0.0);
    END_IF;
    (* Blip court : arme sur le meme front MECANIQUE. Ses propres bascules electriques ne
       peuvent donc jamais le rearmer — meme protection que l'episode d'intermittence. *)
    IF (BlipTransitions > 0) AND (BlipDurationS > 0.0) THEN
        BlipRunning := TRUE;
        BlipTimerS := 0.0;
        BlipCount := 0;
        BlipActive := TRUE;
        (* Ecretage : au-dela de ce plafond, un compteur UDINT pourrait reboucler et rendre
           le blip non terminant (revue du 2026-09-20, F9). *)
        BlipTransitions := MIN(BlipTransitions, CST_BlipMaxTransitions);
    END_IF;
END_IF;

IF BlipRunning THEN
    (* Protocole du blip court : (0) la sortie rejoint d'abord l'etat MECANIQUE — le
       comportement nominal reste donc visible ; puis une excursion contradictoire toutes
       les BlipDurationS, donc de largeur BlipDurationS ; enfin la sortie est rendue a
       l'etat mecanique. Nombre d'excursions = BlipTransitions. *)
    BlipTimerS := BlipTimerS + CycleTimeS;
    IF BlipTimerS >= MAX(CycleTimeS, BlipDurationS) THEN
        BlipTimerS := 0.0;
        IF BlipCount = 0 THEN
            IF ElectricalOutput <> RawDetected THEN
                ElectricalOutput := RawDetected;
                TransitionCount := TransitionCount + 1;
            END_IF;
            BlipCount := 1;
        ELSIF BlipCount <= BlipTransitions THEN
            ElectricalOutput := NOT ElectricalOutput;
            TransitionCount := TransitionCount + 1;
            BlipCount := BlipCount + 1;
        ELSE
            BlipRunning := FALSE;
            BlipActive := FALSE;
            IF ElectricalOutput <> RawDetected THEN
                ElectricalOutput := RawDetected;
                TransitionCount := TransitionCount + 1;
            END_IF;
            DelayTimerS := 0.0;
        END_IF;
    END_IF;
ELSIF EpisodeActive THEN
    EpisodeTimerS := EpisodeTimerS + CycleTimeS;
    ToggleTimerS := ToggleTimerS + CycleTimeS;
    IF ToggleTimerS >= EpisodeTogglePeriodS THEN
        ElectricalOutput := NOT ElectricalOutput;
        ToggleTimerS := 0.0;
        TransitionCount := TransitionCount + 1;
    END_IF;
    IF EpisodeTimerS >= IntermittenceDurationS THEN
        EpisodeActive := FALSE;
        IF ElectricalOutput <> EpisodeTarget THEN
            ElectricalOutput := EpisodeTarget;
            TransitionCount := TransitionCount + 1;
        END_IF;
        DelayTimerS := 0.0;
    END_IF;
ELSIF ElectricalOutput <> RawDetected THEN
    DelayTimerS := DelayTimerS + CycleTimeS;
    IF DelayTimerS >= MAX(0.0, ElectricalDelayS) THEN
        ElectricalOutput := RawDetected;
        DelayTimerS := 0.0;
        TransitionCount := TransitionCount + 1;
    END_IF;
ELSE
    DelayTimerS := 0.0;
END_IF;

(* ---- FB_Sim_Safety.st ---- *)
(* ═══════════════════════════════════════════════════════════════
   🧪 FB_Sim_Safety — Simulation de la chaîne d'AU et du contacteur de puissance
   ───────────────────────────────────────────────────────────────
   📥 Enable            : activation de la simulation (SimulationModeActive AND NOT SensorEmergencyStopChainIsReal)
   📥 SimChainOkBit     : bit opérateur — TRUE = simuler la chaîne AU fermée ; FALSE = chaîne ouverte (non simulée)
   📥 PowerCutOff_A     : demande de coupure PLC canal A (TRUE = OK/fermé) — conservé pour interface, non utilisé par SimChainOk
   📥 PowerCutOff_B     : demande de coupure PLC canal B (TRUE = OK/fermé) — conservé pour interface, non utilisé par SimChainOk
   📥 PowerCutOffRequest: requête de coupure métier (PowerCutOffRequest du FB AU) — TRUE = arrêt d'urgence (chaîne ouverte)
   📥 EmergencyArming   : impulsion de réarmement (EmergencyArming_RQ)
   📥 BtnEmergencyStop   : appui coup-de-poing AU (TRUE = boucle ouverte)
   📥 TestCutActive     : test de redondance en cours (canal A ou B coupé par le FB AU)

   📤 SimChainOk        : simulation de la boucle AU (fermée si SimChainOkBit, ouverte sur coup-de-poing/test/coupure)
   📤 SimContactorOk    : simulation du contacteur engagé (PowerContactorEngaged)

   ⚙️ MÉCANISME GRANULAIRE (contrôle opérateur de la chaîne AU) :
      - `SimChainOkBit` pilote la chaîne : FALSE → chaîne OUVERTE (on ne peut pas armer) ;
        TRUE → chaîne FERMÉE (le bouton Armable s'active, on arme, la séquence teste les sorties).
      - Pendant le test de redondance (TestCutActive), la chaîne CLIGNOTE (s'ouvre pendant TEST_A/B,
        se referme pendant RESTORE_A/B) puis revient à 1 — comme en réel.
      - `PowerCutOffRequest` (coupure métier) ouvre la chaîne → ARRÊT D'URGENCE.
      - `BtnEmergencyStop` (coup-de-poing) ouvre la chaîne.
      - Le contacteur ne s'engage QUE pendant l'impulsion d'armement (EmergencyArming), avec une
        temporisation d'engagement (CST_ContactorEngageDelay), puis s'auto-maintient tant que la
        chaîne est saine ; il retombe (CST_ContactorDropDelay) dès que la chaîne s'ouvre.
      - À la ré-entrée en simulation (Enable FALSE→TRUE), SimChainOkBit = FALSE → chaîne OUVERTE et
        contacteur NON engagé (on n'a pas armé) — pas de faux « OK » immédiat.

   🔒 NON-RÉGRESSION ARMEMENT (dépendance circulaire) :
      - La chaîne n'est PAS fermée par défaut : elle est fermée UNIQUEMENT si l'opérateur pose
        `SimChainOkBit`. Elle ne dépend PAS de PowerCutOff_A/B (qui sont dans le cercle) : le
        réarmement après échec de test de redondance (RedundancyTestFailedCause laté → PowerCutOff_A=FALSE)
        reste possible car la chaîne est maintenue fermée par le bit opérateur, pas par le PLC.
      - L'ouverture « PLC coupe un canal » est représentée par TestCutActive (test redondance) et
        PowerCutOffRequest (coupure métier) — jamais par PowerCutOff_A/B seuls.
   ═══════════════════════════════════════════════════════════════
   📄 Doc métier : DOC/AF/AF_Partie-13_Fonction_Simulation_v2.5.md
*)
FUNCTION_BLOCK FB_Sim_Safety
VAR_INPUT
    Enable            : BOOL; // --> [CMD] Activation de la simulation
    SimChainOkBit     : BOOL; // --> [TST] Bit opérateur : TRUE = simuler chaîne AU fermée
    SimPhaseRotationOkBit : BOOL; // --> [TST] Bit opérateur : TRUE = phases réseau OK simulées ; FALSE = défaut rotation de phases injecté
    PowerCutOff_A     : BOOL; // --> [SAFE] Commande coupure canal A (TRUE = OK/fermé)
    PowerCutOff_B     : BOOL; // --> [SAFE] Commande coupure canal B (TRUE = OK/fermé)
    PowerCutOffRequest: BOOL; // --> [SAFE] Requête coupure métier (TRUE = arrêt d'urgence)
    EmergencyArming   : BOOL; // --> [CMD] Impulsion de réarmement (TRUE = pulse)
    BtnEmergencyStop   : BOOL; // --> [HW] Force l'ouverture de la boucle (TRUE = bouton appuyé/défaut)
    TestCutActive      : BOOL; // --> [SAFE] Test de redondance en cours (canal A ou B coupé par le FB AU)
END_VAR
VAR_OUTPUT
    SimChainOk      : BOOL; // <-- [STAT] Boucle AU simulée saine
    SimContactorOk  : BOOL; // <-- [STAT] Contacteur simulé engagé
    SimPhaseRotationOk : BOOL; // <-- [STAT] Contrôleur de phases simulé : TRUE = phases saines (aucun défaut)
END_VAR
VAR
    ContactorLatch  : BOOL; // . [LOC] Mémorisation de l'auto-maintien du contacteur
    ChainOpenReq    : BOOL; // . [LOC] Demande brute d'ouverture de la chaîne (bit off / coup-de-poing / test / coupure)
    ChainOpen       : BOOL; // . [LOC] État latche de la chaîne (TRUE = ouverte)
    ContactorEngageReq : BOOL; // . [LOC] Demande d'engagement du contacteur (pulse ET chaîne saine)
    TonChainOpen    : TON;  // . [LOC] Temporisation d'ouverture de la chaîne (retombée relais)
    TonChainClose   : TON;  // . [LOC] Temporisation de fermeture de la chaîne (retombée relais)
    TonContactorEngage : TON; // . [LOC] Temporisation d'engagement du contacteur (temps de collage bobine)
    TonContactorDrop   : TON; // . [LOC] Temporisation de retombée du contacteur (temps de décollage bobine)
END_VAR
VAR CONSTANT
    // === TEMPORISATIONS PHYSIQUES SIMULÉES (compatibles séquence FB AU) ===
    // ⚠️ Doivent rester < durées de la séquence FB AU (CST_TestDuration=200ms, CST_ArmingPulseDuration=1s,
    //    CST_ArmingConfirmTimeout=2s) pour que le test de redondance et la confirmation contacteur
    //    restent validés : ouverture/fermeture chaîne < 200ms, engagement contacteur < 1s.
    CST_ChainOpenDelay       : TIME := T#50ms;  // Temps de retombée relais AU (ouverture chaîne)
    CST_ChainCloseDelay      : TIME := T#50ms;  // Temps de retombée relais AU (fermeture chaîne)
    CST_ContactorEngageDelay : TIME := T#100ms; // Temps de collage bobine contacteur (engagement)
    CST_ContactorDropDelay   : TIME := T#50ms;  // Temps de décollage bobine contacteur (retombée)
END_VAR

// === IMPLEMENTATION ===
{region "§1 Gate"}
IF NOT Enable THEN
    SimChainOk     := FALSE;
    SimContactorOk := FALSE;
    SimPhaseRotationOk := FALSE;
    ContactorLatch := FALSE;
    ChainOpen      := TRUE; // Chaîne ouverte par défaut à la ré-entrée (on n'a pas armé)
    ChainOpenReq   := FALSE;
    ContactorEngageReq := FALSE;
    TonChainOpen(IN := FALSE);
    TonChainClose(IN := FALSE);
    TonContactorEngage(IN := FALSE);
    TonContactorDrop(IN := FALSE);
    RETURN;
END_IF;
{endregion}

{region "§2 Chaîne AU (contrôle granulaire + dynamique)"}
// 1. La chaîne AU est saine si l'opérateur la simule fermée (SimChainOkBit = TRUE) ET si aucun
//    événement ne l'ouvre : coup-de-poing (BtnEmergencyStop), test de redondance (TestCutActive),
//    coupure métier (PowerCutOffRequest).
// 🔧 DEADLOCK SIMULATION (corrigé) : la chaîne n'est PAS fermée par défaut ni dépendante de
//    PowerCutOff_A/B (qui sont dans le cercle). Elle est fermée UNIQUEMENT par le bit opérateur
//    `SimChainOkBit`. Le réarmement après échec de test de redondance (RedundancyTestFailedCause laté
//    → PowerCutOff_A=FALSE) reste possible car la chaîne est maintenue fermée par le bit, pas par
//    le PLC. Hors simulation (Enable=FALSE), la chaîne reste pilotée par le matériel via le repli
//    HwReal (PRG_02 §1/§2) — aucune régression sécurité réelle.
// 🆕 DYNAMIQUE : l'ouverture/fermeture suit une temporisation (CST_ChainOpenDelay / CST_ChainCloseDelay)
//    qui simule le temps de retombée des relais AU, tout en restant < 200ms (CST_TestDuration) pour
//    ne pas fausser le test de redondance. Pendant le test, la chaîne clignote (s'ouvre en TEST_A/B,
//    se referme en RESTORE_A/B) puis revient à 1.
ChainOpenReq := (NOT SimChainOkBit) OR BtnEmergencyStop OR TestCutActive OR PowerCutOffRequest;

// Temporisation d'ouverture : la chaîne s'ouvre après CST_ChainOpenDelay de demande soutenue
TonChainOpen(IN := ChainOpenReq, PT := CST_ChainOpenDelay);
// Temporisation de fermeture : la chaîne se ferme après CST_ChainCloseDelay d'absence de demande
TonChainClose(IN := NOT ChainOpenReq, PT := CST_ChainCloseDelay);

// Latch de la chaîne avec temporisations (défaut = ouverte à la ré-entrée)
IF ChainOpenReq THEN
    IF TonChainOpen.Q THEN
        ChainOpen := TRUE;
    END_IF;
ELSE
    IF TonChainClose.Q THEN
        ChainOpen := FALSE;
    END_IF;
END_IF;

SimChainOk := NOT ChainOpen;
{endregion}

{region "§3 Auto-maintien contacteur (dynamique réaliste)"}
// 2. Logique d'auto-maintien (latch) du contacteur avec priorité à la coupure.
// 🆕 DYNAMIQUE : le contacteur ne s'engage QUE pendant l'impulsion d'armement (EmergencyArming)
//    tant que la chaîne est saine, après CST_ContactorEngageDelay (temps de collage bobine), puis
//    s'auto-maintient. Il retombe après CST_ContactorDropDelay (temps de décollage bobine) dès que
//    la chaîne s'ouvre — comme une bobine réelle qui décolle sans alimentation. Ces temporisations
//    restent < CST_ArmingPulseDuration (1s) et CST_ArmingConfirmTimeout (2s) pour que la
//    confirmation contacteur reste validée. À la ré-entrée en simulation, le contacteur est NON
//    engagé (on n'a pas armé).
ContactorEngageReq := EmergencyArming AND SimChainOk;

// Temporisation d'engagement : le contacteur se colle après CST_ContactorEngageDelay de pulse soutenu
TonContactorEngage(IN := ContactorEngageReq, PT := CST_ContactorEngageDelay);
// Temporisation de retombée : le contacteur décolle après CST_ContactorDropDelay de chaîne ouverte
TonContactorDrop(IN := NOT SimChainOk, PT := CST_ContactorDropDelay);

// Latch du contacteur avec priorité à la coupure (retombée > engagement)
IF NOT SimChainOk THEN
    IF TonContactorDrop.Q THEN
        ContactorLatch := FALSE;
    END_IF;
ELSIF ContactorEngageReq THEN
    IF TonContactorEngage.Q THEN
        ContactorLatch := TRUE;
    END_IF;
END_IF;

// Recopie vers la sortie
SimContactorOk := ContactorLatch;

// Contrôleur de phases : simple propagation du bit opérateur (TRUE = sain).
// Inopérant hors simulation (le banc ne publie l'image machine que sous Enable).
SimPhaseRotationOk := SimPhaseRotationOkBit;
{endregion}

(* ---- FB_Sim_SuspendedLoad.st ---- *)
(* DOC: DOC/AF/AF_Partie-13_Fonction_Simulation_v2.5.md
   Pendule reduit : reaction sur chariot sans injection DI directe. *)
FUNCTION_BLOCK PUBLIC FB_Sim_SuspendedLoad
VAR_INPUT
    Enable : BOOL;
    BrakeMechanicallyOpen : BOOL;
    CartAcceleration_Mps2 : REAL;
    Length_M : REAL := 1.5;
    Damping : REAL := 0.35;
    ReactionGain_Mps2 : REAL := 0.20;
    CycleTime_S : REAL := 0.01;
END_VAR
VAR_OUTPUT
    Ready : BOOL;
    Angle_Rad : REAL;
    AngularVelocity_RadPerS : REAL;
    VelocityReaction_Mps : REAL;
END_VAR
VAR
    AngularAccel_RadPerS2 : REAL;
END_VAR
VAR CONSTANT
    CST_Gravity_Mps2 : REAL := 9.81;
    CST_MinLength_M : REAL := 0.1;
    CST_MaxAngle_Rad : REAL := 0.6;
    CST_MaxAngularVelocity_RadPerS : REAL := 4.0;
END_VAR

IF NOT Enable THEN
    Ready := FALSE;
    Angle_Rad := 0.0;
    AngularVelocity_RadPerS := 0.0;
    VelocityReaction_Mps := 0.0;
    RETURN;
END_IF;

VelocityReaction_Mps := 0.0;
IF Length_M > CST_MinLength_M THEN
    AngularAccel_RadPerS2 := -(CST_Gravity_Mps2 / Length_M) * Angle_Rad
        - MAX(0.0, Damping) * AngularVelocity_RadPerS
        - CartAcceleration_Mps2 / Length_M;
    AngularVelocity_RadPerS := LIMIT(-CST_MaxAngularVelocity_RadPerS,
        AngularVelocity_RadPerS + AngularAccel_RadPerS2 * CycleTime_S, CST_MaxAngularVelocity_RadPerS);
    Angle_Rad := LIMIT(-CST_MaxAngle_Rad, Angle_Rad + AngularVelocity_RadPerS * CycleTime_S,
        CST_MaxAngle_Rad);
    IF BrakeMechanicallyOpen THEN
        VelocityReaction_Mps := ReactionGain_Mps2 * Angle_Rad * CycleTime_S;
    END_IF;
END_IF;
Ready := TRUE;

(* ---- FB_Sim_Translation.st ---- *)
(* DOC: DOC/AF/AF_Partie-13_Fonction_Simulation_v2.5.md
   Modele dynamique M3 confine au SimBench. *)
FUNCTION_BLOCK PUBLIC FB_Sim_Translation
VAR_INPUT
    Enable : BOOL;
    ReqTremie : BOOL;
    ReqMaintenance : BOOL;
    SpeedTgt_Pct : REAL;
    (* T301/L1 — SOURCE UNIQUE : le banc ne porte AUCUNE position ni echelle propre.
       Positions capteurs = reglages machine (GVL_PERSISTENT._TranslationPos*_M) et gain =
       gain EFFECTIVEMENT consomme par l'estimateur (PRG_05 FB_Translation_OdometryGain.GainActive),
       passes par PRG_02 -> FB_SimBench. Vitesse chariot = sens x gain x frequence.
       Historique : l'ancienne echelle en dur (30 m / FullTravelTimeS / 40 Hz) a diverge du gain
       reel (T360/T361, sauts de 4 a 9 m) — doublon supprime, gate G518 anti-retour. *)
    PosTremie_M        : REAL := 0.0;   (* --> [CFG] Position capteur Tremie (m) *)
    PosPV_M            : REAL := 1.5;   (* --> [CFG] Position capteur PV (m) *)
    PosP2_M            : REAL := 3.5;   (* --> [CFG] Position capteur P2 (m) *)
    PosP1_M            : REAL := 5.0;   (* --> [CFG] Position capteur P1 (m) *)
    PosMaintenance_M   : REAL := 10.0;  (* --> [CFG] Position capteur Maintenance (m) *)
    GainMetersPerHzSec : REAL := 0.02;  (* --> [CFG] Gain odometrique effectif, m/(Hz.s) *)
    (* Distance capteur extreme -> butee mecanique (seule donnee propre au banc : physique du rail).
       Bornee a CST_MinEndStopMargin_M pour que le capteur extreme reste franchissable. *)
    EndStopMargin_M    : REAL := 0.5;
    BrakeReleaseCmd : BOOL := TRUE;
    (* ECHELLE DE LA CONSIGNE. PRG_02 envoie SpeedCmd_Pct = f / 50 Hz x 100 : le simulateur reconvertit
       avec le MEME maximum, sinon 20 Hz reels (40 %) deviendraient 16 Hz simules.
       Maximum = GVL_PERSISTENT._TranslationMaxFreq_Hz (50 Hz), passe par FB_SimBench (CST_M3MaxFreq_Hz,
       egalite verifiee par G518). Ne pas confondre avec l'ancienne echelle (40 Hz) : echelle
       ODOMETRIQUE (gain 0,02 m/(Hz.s)). *)
    MaxFreq_Hz : REAL := 50.0;
    (* ACCELERATION DU BANC (confort d'essai). Le chariot avance SpeedFactor fois plus vite ET la
       frequence RETOURNEE au PLC est multipliee d'autant : l'estimateur (f x gain) suit exactement
       le chariot, sans saut de recalage, et le ratio publie reste 0,02 m/(Hz.s) (G518).
       Borne 1..5. 1,0 = dynamique reelle. Le frein et la memoire de sens restent sur la frequence
       physique du variateur simule. *)
    SpeedFactor : REAL := 1.0;
    AccelRate_HzPerS : REAL := 20.0;
    DecelRate_HzPerS : REAL := 25.0; // pente d'arret relevee sur trace reelle (rampe variateur / rampe PLC)
    DriveTimeConstantS : REAL := 0.15;
    BrakeOpenDelayS : REAL := 0.10;
    BrakeCloseDelayS : REAL := 0.09;
    BrakeContactDelayS : REAL := 0.01;
    (* FAUTE EXPLICITE frein M3 — defaut FALSE : reproduit le defaut terrain « frein ferme
       alors que le variateur retourne encore 10,00 Hz » (trace 2026-09-04, 26,437 s,
       State.ErrorId=64). La garde nominale 0,5 Hz du frein n'est pas modifiee. *)
    BrakeFaultCloseWhileRunning : BOOL := FALSE;
    BrakeFaultCloseDelay_S : REAL := 0.0;
    (* L3 — FREIN PHYSIQUE (2026-10-28). FALSE = historique (frein ne retombe que sous 0,5 Hz,
       arret instantane). TRUE = frein a manque de courant reel : retombe CloseDelay apres la
       coupure bobine QUELLE QUE SOIT la vitesse, puis le chariot decelere sur le frein
       (BrakeDecel_Mps2) ; frein serre = chariot bloque meme si le variateur pousse. *)
    BrakePhysicalActive : BOOL := FALSE; (* defaut FB = historique ; GVL_Simulation.SimM3BrakePhysicalActive = TRUE (source unique) *)
    BrakeDecel_Mps2 : REAL := 2.0;   (* HYPOTHESE : 0,4 m/s (20 Hz) -> arret ~0,2 s / ~4 cm *)
    (* L4 — CHARIOT LIBRE (2026-10-28). FALSE = historique (chariot esclave de la frequence).
       TRUE = quand le frein est OUVERT et que le variateur n'applique plus de couple (mot a 0
       et rampe variateur terminee), le chariot n'est plus tenu : il garde sa vitesse et subit
       la poussee de la benne suspendue (rapport de masse x g x angle), la pente et le
       frottement de roulement. Valeurs = HYPOTHESES, sans mesure terrain. *)
    CartFreeActive : BOOL := FALSE;
    LoadMassRatio : REAL := 0.5;          (* masse benne / masse totale chariot+benne *)
    RollingFriction_Mps2 : REAL := 0.30;  (* FEM 1.001 : frottement global galets + reducteur accouple *)
    StaticFriction_Mps2 : REAL := 0.35;   (* Seuil de decollement statique (anti-pompage pendulaire) *)
    Slope_Mps2 : REAL := 0.0;             (* composante de pente, + vers Maintenance *)
    (* L5 — came capteurs (vu -> perdu -> retrouve -> fixe), appliquee aux 5 capteurs. *)
    SensorCamDropoutActive : BOOL := FALSE;
    SensorCamDropoutStart_M : REAL := 0.02;
    SensorCamDropoutWidth_M : REAL := 0.04;
    SuspendedLoadLength_M : REAL := 1.5;
    SuspendedLoadDamping : REAL := 0.35;
    LoadReactionGain_Mps2 : REAL := 0.20;
    (* BUTEE MECANIQUE — recul borne apres arret serre.
       0.0 (defaut) conserve EXACTEMENT le comportement historique : position ET vitesse
       figees a la butee (decision de review tracee, correctif « contact rigide »).
       > 0 : l'inertie du chariot reste absorbee par la butee, MAIS la reaction de la charge
       peut ressortir le chariot de la zone capteur — comportement observe sur la trace
       terrain du 2026-09-04 a 26,437 s (Tremie actif 1 echantillon puis perdu
       definitivement). Valeur SYNTHETIQUE, en attente de mesure terrain. *)
    EndStopRecoilMax_M : REAL := 0.0;
    LoadFrequencyDroopGain_Hz : REAL := 0.50;
    SensorJitterAmplitude_M : REAL := 0.01;
    SensorStabilizationS : REAL := 1.0;
    SensorElectricalDelayS : REAL := 0.01;
    SensorIntermittenceActive : BOOL := FALSE;
    SensorLoadAngleTriggerRad : REAL := 0.01;
    SensorScenarioSeed : UDINT := 3001;
    SensorHysteresis_M : REAL := 0.02;
    SensorIntermittencePeriodS : REAL := 0.12;
    (* BLIP COURT — second profil capteur, independant du train ~1 s ci-dessus.
       BlipTransitions = 0 (defaut) : profil historique strictement inchange.
       Valeurs de trace : Tremie 1 excursion de 0,2 s (2 echantillons a 100 ms),
       PV 1 excursion de 0,1 s (1 echantillon).
       ⚠️ LIMITE CONNUE (revue 2026-09-20, F11) : UNE SEULE largeur globale est appliquee aux
       cinq capteurs. Les deux signatures de la trace (Tremie 0,200 s et PV 0,100 s) ne sont
       donc PAS rejouables dans la meme passe : il faut deux executions avec des valeurs
       differentes de SensorBlipDurationS. Une largeur par capteur exigerait un
       ARRAY[1..5] OF REAL, non retenu dans ce lot. *)
    SensorBlipTransitions : UDINT := 0;
    SensorBlipDurationS : REAL := 0.2;
END_VAR
VAR_OUTPUT
    PosTremie : BOOL;
    PosPV : BOOL;
    PosP2 : BOOL;
    PosP1 : BOOL;
    PosMaintenance : BOOL;
    FrequencyCmd_Hz : REAL;
    ElectricalFrequency_Hz : REAL;
    ActualFrequency_Hz : REAL;
    BrakeCoilEnergized : BOOL;
    BrakeMechanicallyOpen : BOOL;
    BrakeContactOpen : BOOL;
    BrakeFaultCloseActive : BOOL;
    PositionTrue_M : REAL;
    VelocityTrue_Mps : REAL;
    LoadAngle_Rad : REAL;
    SensorPosition_M : REAL;
    SensorTransitionCount : UDINT;
    SensorBlipActive : BOOL;
    HardStopTremieActive : BOOL;
    HardStopMaintenanceActive : BOOL;
    (* L2 — OBSERVATION (aucun effet sur le modele ni sur le programme) *)
    ObsOvershootLast_M : REAL;          (* Distance roulee entre le 1er front du dernier capteur d'arret (Tremie, P1, Maintenance) et l'arret *)
    ObsOvershootSensorId : INT;         (* 1 = Tremie, 3 = P1, 5 = Maintenance, 0 = aucun *)
    ObsEndStopHitCount : UDINT;         (* Nombre de chocs en butee mecanique *)
    ObsEndStopImpactSpeed_Mps : REAL;   (* Vitesse au dernier choc en butee *)
    ObsBrakeClosedMovingCount : UDINT;  (* Nombre de fermetures mecaniques du frein chariot en mouvement *)
    ObsCartFree : BOOL;                 (* L4 : frein ouvert ET variateur sans couple -> chariot libre *)
    ObsFreeRollLast_M : REAL;           (* L4 : distance parcourue pendant le dernier episode libre *)
END_VAR
VAR
    ObsArmed : BOOL;                    (* Front capteur d'arret vu, arret pas encore constate *)
    ObsEdgePosition_M : REAL;           (* Position vraie au 1er front du capteur d'arret *)
    ObsPrevTremie : BOOL;
    ObsPrevP1 : BOOL;
    ObsPrevMaintenance : BOOL;
    ObsPrevBrakeOpen : BOOL;
    ObsPrevHardStop : BOOL;
    ObsSpeedBeforeStop_Mps : REAL;      (* Vitesse du scan avant le calcul de butee *)
    DriveTorqueActive : BOOL;           (* L4 : variateur commande ou encore en rampe -> chariot tenu *)
    FreeAccel_Mps2 : REAL;              (* L4 : acceleration nette du chariot libre *)
    FreeVelocity_Mps : REAL;           (* Vitesse apres integration de la force externe *)
    FrictionStep_Mps : REAL;           (* Impulsion dissipative maximale sur le pas *)
    FreeRollStart_M : REAL;             (* L4 : position au debut de l'episode libre *)
    instCycleTime : FB_CycleTime;
    Initialized : BOOL;
    DirectionSign : REAL;
    (* Sens de deplacement MEMORISE. La commande peut etre retiree AVANT l'arret physique
       (deceleration libre du variateur) : le sens du dernier ordre valide est conserve tant
       que le variateur retourne de la vitesse, puis purge a l'arret. Sans cette memoire, la
       vitesse du chariot s'effondrait au scan de retrait de commande alors que la frequence
       retournee decroit encore.
       ⚠️ ORDRE DE GRANDEUR NON MESURE : la trace terrain ne contient AUCUNE variable de
       position (15 TraceVariable : DI, frequences, mots d'etat, erreurs). La distance de
       roue libre de la fenetre 14,67 -> 16,16 s est donc une ESTIMATION dependante du modele
       d'echelle, qui vaut approximativement 1,1 a 1,3 m selon la methode d'integration
       retenue (gain audit 0,0551 m/(Hz.s)). A ne pas citer comme une mesure. *)
    TravelDirection : REAL;
    FrequencyTarget_Hz : REAL;
    SpeedFactorApplied : REAL := 1.0;
    CycleTimeS : REAL;
    EndStopTremie_M : REAL;       (* butee mecanique cote Tremie = capteur Tremie - marge *)
    EndStopMaintenance_M : REAL;  (* butee mecanique cote Maintenance = capteur Maintenance + marge *)
    VelocityTarget_Mps : REAL;
    CartAcceleration_Mps2 : REAL;
    PreviousVelocity_Mps : REAL;
    PositionCandidate_M : REAL;
    (* Recul de butee ECRETE a la course : une valeur d'entree aberrante ne peut pas
       autoriser une position hors des butees (revue du 2026-09-20, F8). *)
    RecoilMax_M : REAL;
    SensorNoiseState : REAL := 0.371;
    SensorNoise_M : REAL;
    instSensorTremie : FB_Sim_PositionSensor;
    instSensorPV : FB_Sim_PositionSensor;
    instSensorP2 : FB_Sim_PositionSensor;
    instSensorP1 : FB_Sim_PositionSensor;
    instSensorMaintenance : FB_Sim_PositionSensor;
    instDrive : FB_Sim_TranslationDrive;
    instBrake : FB_Sim_TranslationBrake;
    instSuspendedLoad : FB_Sim_SuspendedLoad;
END_VAR
VAR CONSTANT
    (* Marge mini capteur extreme -> butee : au-dela de l'hysteresis capteur, sinon le mot
       11111 / 00000 ne pourrait jamais etre produit (capteur colle a la butee). *)
    CST_MinEndStopMargin_M : REAL := 0.05;
    (* Meme seuil d'arret que FB_Sim_TranslationBrake.CST_StopFrequency_Hz (0,5 Hz).
       Valide par la trace terrain du 2026-09-04 : frein ouvert a 0,60 Hz, ferme a 0,00 Hz. *)
    CST_StopFrequency_Hz : REAL := 0.5;
END_VAR

instCycleTime(DefaultValueS := 0.010);
(* Le modele mono-pas suit le temps de cycle reel jusqu'a 100 ms. Cette borne
   evite de ralentir artificiellement la dynamique lorsque la trace est executee
   dans VISU_TASK (environ 100 ms), tout en restant stable pour le pendule reduit.
   Au-dela, FB_CycleTime fournit deja son temps de secours et aucun saut aberrant
   n'est accepte. La qualification des delais sub-100 ms exige toutefois une tache
   de trace plus rapide que 100 ms. *)
CycleTimeS := LIMIT(0.001, instCycleTime.CycleTimeS, 0.100);

(* Butees mecaniques derivees des capteurs extremes (reglages machine) + marge du rail. *)
EndStopTremie_M := PosTremie_M - MAX(EndStopMargin_M, CST_MinEndStopMargin_M);
EndStopMaintenance_M := PosMaintenance_M + MAX(EndStopMargin_M, CST_MinEndStopMargin_M);

IF NOT Enable THEN
    Initialized := FALSE;
    instDrive(Enable := FALSE);
    instBrake(Enable := FALSE);
    instSuspendedLoad(Enable := FALSE);
    FrequencyCmd_Hz := 0.0;
    ElectricalFrequency_Hz := 0.0;
    ActualFrequency_Hz := 0.0;
    BrakeMechanicallyOpen := FALSE;
    BrakeContactOpen := FALSE;
    BrakeCoilEnergized := FALSE;
    BrakeFaultCloseActive := FALSE;
    PositionTrue_M := PosP1_M;
    VelocityTrue_Mps := 0.0;
    PreviousVelocity_Mps := 0.0;
    TravelDirection := 0.0;
    LoadAngle_Rad := 0.0;
    SensorTransitionCount := 0;
    SensorBlipActive := FALSE;
    HardStopTremieActive := FALSE;
    HardStopMaintenanceActive := FALSE;
    (* Repli deterministe compatible avec le mot thermometre P1 = 00011. *)
    PosTremie := FALSE;
    PosPV := FALSE;
    PosP2 := FALSE;
    PosP1 := TRUE;
    PosMaintenance := TRUE;
    instSensorTremie(Enable := FALSE);
    instSensorPV(Enable := FALSE);
    instSensorP2(Enable := FALSE);
    instSensorP1(Enable := FALSE);
    instSensorMaintenance(Enable := FALSE);
    RETURN;
ELSIF NOT Initialized THEN
    Initialized := TRUE;
    PositionTrue_M := PosP1_M;
    TravelDirection := 0.0;
END_IF;

IF Enable THEN
    DirectionSign := 0.0;
    IF ReqTremie AND NOT ReqMaintenance THEN
        DirectionSign := -1.0;
    ELSIF ReqMaintenance AND NOT ReqTremie THEN
        DirectionSign := 1.0;
    END_IF;

    FrequencyTarget_Hz := LIMIT(0.0, ABS(SpeedTgt_Pct) * MaxFreq_Hz / 100.0, MaxFreq_Hz);
    IF DirectionSign = 0.0 THEN
        FrequencyTarget_Hz := 0.0;
    END_IF;
    instDrive(Enable := TRUE, FrequencyTgt_Hz := FrequencyTarget_Hz,
        AccelRate_HzPerS := AccelRate_HzPerS, DecelRate_HzPerS := DecelRate_HzPerS,
        TimeConstant_S := DriveTimeConstantS,
        LoadAngularVelocity_RadPerS := instSuspendedLoad.AngularVelocity_RadPerS,
        LoadFrequencyDroopGain_Hz := LoadFrequencyDroopGain_Hz, CycleTime_S := CycleTimeS);
    FrequencyCmd_Hz := instDrive.FrequencyCmd_Hz;
    ElectricalFrequency_Hz := instDrive.ElectricalFrequency_Hz;
    SpeedFactorApplied := LIMIT(1.0, SpeedFactor, 5.0);
    ActualFrequency_Hz := instDrive.ActualFrequency_Hz * SpeedFactorApplied;
    instBrake(Enable := TRUE, ReleaseCmd := BrakeReleaseCmd,
        ActualFrequency_Hz := instDrive.ActualFrequency_Hz, OpenDelay_S := BrakeOpenDelayS,
        CloseDelay_S := BrakeCloseDelayS, ContactDelay_S := BrakeContactDelayS,
        CycleTime_S := CycleTimeS,
        FaultCloseWhileRunning := BrakeFaultCloseWhileRunning,
        FaultCloseDelay_S := BrakeFaultCloseDelay_S,
        PhysicalBrakeActive := BrakePhysicalActive);
    BrakeCoilEnergized := instBrake.CoilEnergized;
    BrakeMechanicallyOpen := instBrake.MechanicallyOpen;
    BrakeContactOpen := instBrake.ContactOpen;
    BrakeFaultCloseActive := instBrake.FaultCloseActive;

    (* Sens memorise (C3). Regles, dans cet ordre :
       1. un ordre simple valide (re)memorise le sens ;
       2. deux ordres contradictoires neutralisent immediatement le sens — aucune
          excitation inventee (preserve TC-T300-MEC-030) ;
       3. commande retiree : le sens est CONSERVE tant que le variateur retourne de la
          vitesse (deceleration libre), puis purge des que la vitesse est nulle. *)
    IF ReqTremie AND NOT ReqMaintenance THEN
        TravelDirection := -1.0;
    ELSIF ReqMaintenance AND NOT ReqTremie THEN
        TravelDirection := 1.0;
    ELSIF ReqTremie AND ReqMaintenance THEN
        TravelDirection := 0.0;
    ELSIF ABS(instDrive.ActualFrequency_Hz) <= CST_StopFrequency_Hz THEN
        TravelDirection := 0.0;
    END_IF;

    PreviousVelocity_Mps := VelocityTrue_Mps;
    IF BrakeMechanicallyOpen THEN
        (* Source unique : meme gain que l'estimateur machine (vitesse = gain x frequence). *)
        VelocityTarget_Mps := TravelDirection * MAX(0.0, GainMetersPerHzSec) * ActualFrequency_Hz;
    ELSE
        VelocityTarget_Mps := 0.0;
    END_IF;
    (* L4 : le variateur tient le chariot tant qu'il est commande ou que sa SORTIE electrique
       alimente encore le moteur (rampe + reponse) ; ensuite, plus aucun couple.
       Reprise de commande en roue libre : pas de reprise a la volee (le variateur repart de 0 Hz). *)
    DriveTorqueActive := (DirectionSign <> 0.0) OR (instDrive.ElectricalFrequency_Hz > CST_StopFrequency_Hz);
    ObsCartFree := CartFreeActive AND BrakeMechanicallyOpen AND NOT DriveTorqueActive;
    IF ObsCartFree THEN
        (* Poussee de la benne (angle du scan precedent) + pente - frottement oppose au mouvement. *)
        (* Pendule sur chariot libre : x'' = m_benne / m_chariot x g x theta = r / (1 - r) x g x theta. *)
        FreeAccel_Mps2 := (LIMIT(0.0, LoadMassRatio, 0.9) / (1.0 - LIMIT(0.0, LoadMassRatio, 0.9)))
                          * 9.81 * instSuspendedLoad.Angle_Rad + Slope_Mps2;
        IF ABS(VelocityTrue_Mps) < 0.001 THEN
            (* Adherence statique au repos : ne decolle que si la poussee depasse le frottement statique *)
            IF ABS(FreeAccel_Mps2) <= MAX(0.0, StaticFriction_Mps2) THEN
                FreeAccel_Mps2 := 0.0;
                VelocityTrue_Mps := 0.0;
            ELSIF FreeAccel_Mps2 > 0.0 THEN
                FreeAccel_Mps2 := FreeAccel_Mps2 - MAX(0.0, StaticFriction_Mps2);
            ELSE
                FreeAccel_Mps2 := FreeAccel_Mps2 + MAX(0.0, StaticFriction_Mps2);
            END_IF;
            VelocityTrue_Mps := VelocityTrue_Mps + FreeAccel_Mps2 * CycleTimeS;
        ELSE
            (* La force externe peut inverser le mouvement ; le frottement ne peut
               que reduire sa vitesse, au plus jusqu'a zero. *)
            FreeVelocity_Mps := VelocityTrue_Mps + FreeAccel_Mps2 * CycleTimeS;
            FrictionStep_Mps := MAX(0.0, RollingFriction_Mps2) * CycleTimeS;
            IF (((VelocityTrue_Mps > 0.0) AND (FreeVelocity_Mps <= 0.0))
                OR ((VelocityTrue_Mps < 0.0) AND (FreeVelocity_Mps >= 0.0)))
                AND (ABS(FreeAccel_Mps2) <= MAX(0.0, StaticFriction_Mps2)) THEN
                (* Passage par zero pendant le pas : l'adherence interdit un redemarrage
                   sous le seuil statique, meme si la force est opposee au mouvement. *)
                VelocityTrue_Mps := 0.0;
            ELSIF FreeVelocity_Mps > 0.0 THEN
                VelocityTrue_Mps := MAX(0.0, FreeVelocity_Mps - FrictionStep_Mps);
            ELSE
                VelocityTrue_Mps := MIN(0.0, FreeVelocity_Mps + FrictionStep_Mps);
            END_IF;
        END_IF;
    ELSIF BrakeMechanicallyOpen THEN
        (* Vitesse suivant directement le variateur (deja filtre par instDrive) sans double PT1 *)
        VelocityTrue_Mps := VelocityTarget_Mps;
    ELSIF BrakePhysicalActive THEN
        (* L3 : frein serre -> deceleration sur le frein jusqu'a l'arret, puis chariot bloque. *)
        IF VelocityTrue_Mps > 0.0 THEN
            VelocityTrue_Mps := MAX(0.0, VelocityTrue_Mps - MAX(0.0, BrakeDecel_Mps2) * CycleTimeS);
        ELSE
            VelocityTrue_Mps := MIN(0.0, VelocityTrue_Mps + MAX(0.0, BrakeDecel_Mps2) * CycleTimeS);
        END_IF;
    ELSE
        VelocityTrue_Mps := 0.0;   (* historique : arret instantane *)
    END_IF;
    ObsSpeedBeforeStop_Mps := VelocityTrue_Mps;
    HardStopTremieActive := FALSE;
    HardStopMaintenanceActive := FALSE;
    PositionCandidate_M := PositionTrue_M + VelocityTrue_Mps * CycleTimeS;
    IF PositionCandidate_M < EndStopTremie_M THEN
        PositionTrue_M := EndStopTremie_M;
        VelocityTrue_Mps := 0.0;
        HardStopTremieActive := TRUE;
    ELSIF PositionCandidate_M > EndStopMaintenance_M THEN
        PositionTrue_M := EndStopMaintenance_M;
        VelocityTrue_Mps := 0.0;
        HardStopMaintenanceActive := TRUE;
    END_IF;
    CartAcceleration_Mps2 := (VelocityTrue_Mps - PreviousVelocity_Mps) / CycleTimeS;
    instSuspendedLoad(Enable := TRUE, BrakeMechanicallyOpen := BrakeMechanicallyOpen,
        CartAcceleration_Mps2 := CartAcceleration_Mps2, Length_M := SuspendedLoadLength_M,
        Damping := SuspendedLoadDamping, ReactionGain_Mps2 := LoadReactionGain_Mps2,
        CycleTime_S := CycleTimeS);
    LoadAngle_Rad := instSuspendedLoad.Angle_Rad;
    IF HardStopTremieActive OR HardStopMaintenanceActive THEN
        RecoilMax_M := MIN(MAX(0.0, EndStopRecoilMax_M), EndStopMaintenance_M - EndStopTremie_M);
        IF (RecoilMax_M > 0.0) AND BrakeMechanicallyOpen THEN
            (* Recul autorise UNIQUEMENT en s'eloignant de la butee touchee, borne par
               EndStopRecoilMax_M : jamais plus loin dans la butee, jamais de saut cache. *)
            VelocityTrue_Mps := VelocityTrue_Mps + instSuspendedLoad.VelocityReaction_Mps;
            (* Contre une butee, l'entrainement DECROCHE : il ne maintient pas une consigne de
               vitesse dans l'obstacle. Sans cette purge, la consigne de vitesse ecrasait en
               permanence la reaction de charge et le chariot ne pouvait jamais ressortir de
               la zone capteur (recul alors impossible, quelle que soit la charge). *)
            TravelDirection := 0.0;
            IF HardStopTremieActive THEN
                VelocityTrue_Mps := MAX(0.0, VelocityTrue_Mps);
                PositionCandidate_M := LIMIT(EndStopTremie_M,
                    PositionTrue_M + VelocityTrue_Mps * CycleTimeS,
                    EndStopTremie_M + RecoilMax_M);
            ELSE
                VelocityTrue_Mps := MIN(0.0, VelocityTrue_Mps);
                PositionCandidate_M := LIMIT(EndStopMaintenance_M - RecoilMax_M,
                    PositionTrue_M + VelocityTrue_Mps * CycleTimeS,
                    EndStopMaintenance_M);
            END_IF;
            PositionTrue_M := PositionCandidate_M;
        ELSE
            VelocityTrue_Mps := 0.0;
        END_IF;
    ELSE
        IF NOT ObsCartFree THEN
            (* Reaction historique (negligeable) ; en mode libre la poussee est deja integree (L4). *)
            VelocityTrue_Mps := VelocityTrue_Mps + instSuspendedLoad.VelocityReaction_Mps;
        END_IF;
        PositionCandidate_M := PositionTrue_M + VelocityTrue_Mps * CycleTimeS;
        IF PositionCandidate_M < EndStopTremie_M THEN
            PositionTrue_M := EndStopTremie_M;
            VelocityTrue_Mps := 0.0;
            HardStopTremieActive := TRUE;
        ELSIF PositionCandidate_M > EndStopMaintenance_M THEN
            PositionTrue_M := EndStopMaintenance_M;
            VelocityTrue_Mps := 0.0;
            HardStopMaintenanceActive := TRUE;
        ELSE
            PositionTrue_M := PositionCandidate_M;
        END_IF;
    END_IF;
END_IF;

IF Enable AND (ABS(LoadAngle_Rad) > 0.0001) THEN
    SensorNoiseState := 3.91 * SensorNoiseState * (1.0 - SensorNoiseState);
    SensorNoise_M := (2.0 * SensorNoiseState - 1.0) * SensorJitterAmplitude_M;
ELSE
    SensorNoise_M := 0.0;
END_IF;
(* Les capteurs sont fixes au rail et observent le chariot. Le balancier agit
   seulement par la reaction mecanique sur PositionTrue_M et conditionne un
   episode electrique ; aucune deflexion de godet n'est injectee directement. *)
SensorPosition_M := PositionTrue_M + SensorNoise_M;
(* Les capteurs M3 sont volontairement cumulatifs : 11111 -> 00000. Chaque
   brique garde son hysteresis et son episode propres ; aucun timer partage ne
   peut masquer un front d'un autre capteur. *)
instSensorTremie(Enable := Enable, Position_M := SensorPosition_M,
    Threshold_M := PosTremie_M, Hysteresis_M := SensorHysteresis_M,
    ElectricalDelayS := SensorElectricalDelayS, IntermittenceActive := SensorIntermittenceActive
        AND (ABS(LoadAngle_Rad) >= SensorLoadAngleTriggerRad),
    IntermittenceDurationS := SensorStabilizationS, IntermittencePeriodS := SensorIntermittencePeriodS,
    ScenarioSeed := SensorScenarioSeed + 11,
    BlipTransitions := SensorBlipTransitions, BlipDurationS := SensorBlipDurationS,
    CamDropoutActive := SensorCamDropoutActive, CamDropoutStart_M := SensorCamDropoutStart_M,
    CamDropoutWidth_M := SensorCamDropoutWidth_M,
    FiniteCamActive := TRUE, CamLength_M := 0.04,
    CycleTimeS := CycleTimeS);
instSensorPV(Enable := Enable, Position_M := SensorPosition_M,
    Threshold_M := PosPV_M, Hysteresis_M := SensorHysteresis_M,
    ElectricalDelayS := SensorElectricalDelayS, IntermittenceActive := SensorIntermittenceActive
        AND (ABS(LoadAngle_Rad) >= SensorLoadAngleTriggerRad),
    IntermittenceDurationS := SensorStabilizationS, IntermittencePeriodS := SensorIntermittencePeriodS,
    ScenarioSeed := SensorScenarioSeed + 23,
    BlipTransitions := SensorBlipTransitions, BlipDurationS := SensorBlipDurationS,
    CamDropoutActive := SensorCamDropoutActive, CamDropoutStart_M := SensorCamDropoutStart_M,
    CamDropoutWidth_M := SensorCamDropoutWidth_M,
    CycleTimeS := CycleTimeS);
instSensorP2(Enable := Enable, Position_M := SensorPosition_M,
    Threshold_M := PosP2_M, Hysteresis_M := SensorHysteresis_M,
    ElectricalDelayS := SensorElectricalDelayS, IntermittenceActive := SensorIntermittenceActive
        AND (ABS(LoadAngle_Rad) >= SensorLoadAngleTriggerRad),
    IntermittenceDurationS := SensorStabilizationS, IntermittencePeriodS := SensorIntermittencePeriodS,
    ScenarioSeed := SensorScenarioSeed + 37,
    BlipTransitions := SensorBlipTransitions, BlipDurationS := SensorBlipDurationS,
    CamDropoutActive := SensorCamDropoutActive, CamDropoutStart_M := SensorCamDropoutStart_M,
    CamDropoutWidth_M := SensorCamDropoutWidth_M,
    CycleTimeS := CycleTimeS);
instSensorP1(Enable := Enable, Position_M := SensorPosition_M,
    Threshold_M := PosP1_M, Hysteresis_M := SensorHysteresis_M,
    ElectricalDelayS := SensorElectricalDelayS, IntermittenceActive := SensorIntermittenceActive
        AND (ABS(LoadAngle_Rad) >= SensorLoadAngleTriggerRad),
    IntermittenceDurationS := SensorStabilizationS, IntermittencePeriodS := SensorIntermittencePeriodS,
    ScenarioSeed := SensorScenarioSeed + 53,
    BlipTransitions := SensorBlipTransitions, BlipDurationS := SensorBlipDurationS,
    CamDropoutActive := SensorCamDropoutActive, CamDropoutStart_M := SensorCamDropoutStart_M,
    CamDropoutWidth_M := SensorCamDropoutWidth_M,
    CycleTimeS := CycleTimeS);
instSensorMaintenance(Enable := Enable, Position_M := SensorPosition_M,
    Threshold_M := PosMaintenance_M, Hysteresis_M := SensorHysteresis_M,
    ElectricalDelayS := SensorElectricalDelayS, IntermittenceActive := SensorIntermittenceActive
        AND (ABS(LoadAngle_Rad) >= SensorLoadAngleTriggerRad),
    IntermittenceDurationS := SensorStabilizationS, IntermittencePeriodS := SensorIntermittencePeriodS,
    ScenarioSeed := SensorScenarioSeed + 71,
    BlipTransitions := SensorBlipTransitions, BlipDurationS := SensorBlipDurationS,
    CamDropoutActive := SensorCamDropoutActive, CamDropoutStart_M := SensorCamDropoutStart_M,
    CamDropoutWidth_M := SensorCamDropoutWidth_M,
    CycleTimeS := CycleTimeS);

PosTremie := instSensorTremie.ElectricalOutput;
PosPV := instSensorPV.ElectricalOutput;
PosP2 := instSensorP2.ElectricalOutput;
PosP1 := instSensorP1.ElectricalOutput;
PosMaintenance := instSensorMaintenance.ElectricalOutput;
SensorTransitionCount := instSensorTremie.TransitionCount + instSensorPV.TransitionCount
    + instSensorP2.TransitionCount + instSensorP1.TransitionCount
    + instSensorMaintenance.TransitionCount;
SensorBlipActive := instSensorTremie.BlipActive OR instSensorPV.BlipActive
    OR instSensorP2.BlipActive OR instSensorP1.BlipActive
    OR instSensorMaintenance.BlipActive;

(* ── L2 OBSERVATION (lecture seule, aucun effet sur le modele) ───────────────────────── *)
IF Enable THEN
    (* Frein serre en mouvement : front de fermeture mecanique avec vitesse non nulle. *)
    IF ObsPrevBrakeOpen AND NOT BrakeMechanicallyOpen AND (ABS(PreviousVelocity_Mps) > 0.03) THEN
        ObsBrakeClosedMovingCount := ObsBrakeClosedMovingCount + 1;
    END_IF;
    ObsPrevBrakeOpen := BrakeMechanicallyOpen;

    (* Choc en butee : front de HardStop, vitesse avant contact. *)
    IF (HardStopTremieActive OR HardStopMaintenanceActive) AND NOT ObsPrevHardStop THEN
        ObsEndStopHitCount := ObsEndStopHitCount + 1;
        ObsEndStopImpactSpeed_Mps := ABS(ObsSpeedBeforeStop_Mps);
    END_IF;
    ObsPrevHardStop := HardStopTremieActive OR HardStopMaintenanceActive;

    (* Depassement : 1er front d'un capteur d'arret (Tremie montant, P1 dans les deux sens,
       Maintenance descendant) -> position memorisee ; les rebonds du MEME capteur sont ignores
       tant que l'arret n'est pas constate ; un autre capteur franchi remplace le repere. *)
    (* Armement seulement chariot en mouvement : un rebond capteur a l'arret n'ecrase pas la mesure. *)
    IF ABS(VelocityTrue_Mps) <= 0.005 THEN
        ObsArmed := ObsArmed;   (* chariot a l'arret : aucun armement *)
    ELSIF (PosTremie AND NOT ObsPrevTremie) AND NOT (ObsArmed AND ObsOvershootSensorId = 1) THEN
        ObsArmed := TRUE; ObsOvershootSensorId := 1; ObsEdgePosition_M := PositionTrue_M;
    ELSIF (PosP1 <> ObsPrevP1) AND NOT (ObsArmed AND ObsOvershootSensorId = 3) THEN
        ObsArmed := TRUE; ObsOvershootSensorId := 3; ObsEdgePosition_M := PositionTrue_M;
    ELSIF (ObsPrevMaintenance AND NOT PosMaintenance) AND NOT (ObsArmed AND ObsOvershootSensorId = 5) THEN
        ObsArmed := TRUE; ObsOvershootSensorId := 5; ObsEdgePosition_M := PositionTrue_M;
    END_IF;
    ObsPrevTremie := PosTremie;
    ObsPrevP1 := PosP1;
    ObsPrevMaintenance := PosMaintenance;

    (* L4 : distance de l'episode libre (frein ouvert, variateur sans couple). *)
    IF NOT ObsCartFree THEN
        FreeRollStart_M := PositionTrue_M;
    ELSE
        ObsFreeRollLast_M := ABS(PositionTrue_M - FreeRollStart_M);
    END_IF;

    IF ObsArmed AND (ABS(VelocityTrue_Mps) < 0.001) THEN
        ObsOvershootLast_M := ABS(PositionTrue_M - ObsEdgePosition_M);
        ObsArmed := FALSE;
    END_IF;
END_IF;

(* ---- FB_Sim_TranslationBrake.st ---- *)
(* DOC: DOC/AF/AF_Partie-13_Fonction_Simulation_v2.5.md
   Chaine bobine, effet mecanique et contact frein M3. *)
FUNCTION_BLOCK PUBLIC FB_Sim_TranslationBrake
VAR_INPUT
    Enable : BOOL;
    ReleaseCmd : BOOL;
    ActualFrequency_Hz : REAL;
    OpenDelay_S : REAL := 0.10;
    CloseDelay_S : REAL := 0.09;
    ContactDelay_S : REAL := 0.01;
    CycleTime_S : REAL := 0.01;
    (* Branche de FAUTE EXPLICITE — defaut FALSE : chemin nominal strictement inchange.
       Rejoue le defaut terrain « cause 6 instantanee » : contact frein ferme alors que le
       variateur retourne encore de la vitesse (trace 2026-09-04, 26,437 s, 10,00 Hz,
       State.ErrorId=64). La garde nominale CST_StopFrequency_Hz est CONSERVEE telle quelle :
       elle est validee par la meme trace (frein ouvert a 0,60 Hz, ferme a 0,00 Hz). *)
    FaultCloseWhileRunning : BOOL := FALSE;
    FaultCloseDelay_S : REAL := 0.0;
    (* L3 — FREIN PHYSIQUE (2026-10-28). FALSE = historique : la retombee mecanique attend
       f <= 0,5 Hz (garde qui recopiait la logique PLC dans l'usine simulee). TRUE = frein a
       manque de courant reel : retombe CloseDelay_S apres la coupure bobine, QUELLE QUE SOIT
       la vitesse. *)
    PhysicalBrakeActive : BOOL := FALSE; (* defaut FB = historique ; la simulation M3 passe TRUE via GVL_Simulation (source unique) *)
END_VAR
VAR_OUTPUT
    Ready : BOOL;
    CoilEnergized : BOOL;
    MechanicallyOpen : BOOL;
    ContactOpen : BOOL;
    FaultCloseActive : BOOL;   (* <-- [DIAG] Branche de faute effectivement appliquee ce scan *)
END_VAR
VAR
    MechanicalTimer_S : REAL;
    ContactTimer_S : REAL;
    FaultTimer_S : REAL;
END_VAR
VAR CONSTANT
    CST_StopFrequency_Hz : REAL := 0.5;
END_VAR

IF NOT Enable THEN
    Ready := FALSE;
    CoilEnergized := FALSE;
    MechanicallyOpen := FALSE;
    ContactOpen := FALSE;
    FaultCloseActive := FALSE;
    MechanicalTimer_S := 0.0;
    ContactTimer_S := 0.0;
    FaultTimer_S := 0.0;
    RETURN;
END_IF;

(* Faute explicite : chronometre propre, remis a zero des que le stimulus retombe. *)
IF FaultCloseWhileRunning THEN
    FaultTimer_S := FaultTimer_S + CycleTime_S;
ELSE
    FaultTimer_S := 0.0;
END_IF;
FaultCloseActive := FaultCloseWhileRunning AND (FaultTimer_S >= MAX(0.0, FaultCloseDelay_S));

(* La faute fait retomber la bobine : l'etat electrique publie reste coherent avec la
   fermeture mecanique observee (jamais « bobine energisee ET frein serre »). *)
CoilEnergized := ReleaseCmd AND NOT FaultCloseActive;
IF CoilEnergized THEN
    IF NOT MechanicallyOpen THEN
        MechanicalTimer_S := MechanicalTimer_S + CycleTime_S;
        IF MechanicalTimer_S >= MAX(0.0, OpenDelay_S) THEN
            MechanicallyOpen := TRUE;
            MechanicalTimer_S := 0.0;
        END_IF;
    ELSE
        MechanicalTimer_S := 0.0;
    END_IF;
ELSIF FaultCloseActive OR PhysicalBrakeActive OR (ActualFrequency_Hz <= CST_StopFrequency_Hz) THEN
    IF MechanicallyOpen THEN
        MechanicalTimer_S := MechanicalTimer_S + CycleTime_S;
        IF MechanicalTimer_S >= MAX(0.0, CloseDelay_S) THEN
            MechanicallyOpen := FALSE;
            MechanicalTimer_S := 0.0;
        END_IF;
    ELSE
        MechanicalTimer_S := 0.0;
    END_IF;
ELSE
    MechanicalTimer_S := 0.0;
END_IF;
IF MechanicallyOpen <> ContactOpen THEN
    ContactTimer_S := ContactTimer_S + CycleTime_S;
    IF ContactTimer_S >= MAX(0.0, ContactDelay_S) THEN
        ContactOpen := MechanicallyOpen;
        ContactTimer_S := 0.0;
    END_IF;
ELSE
    ContactTimer_S := 0.0;
END_IF;
Ready := TRUE;

(* ---- FB_Sim_TranslationDrive.st ---- *)
(* DOC: DOC/AF/AF_Partie-13_Fonction_Simulation_v2.5.md
   Dynamique reduite du variateur M3, sans commande metier. *)
FUNCTION_BLOCK PUBLIC FB_Sim_TranslationDrive
VAR_INPUT
    Enable : BOOL;
    FrequencyTgt_Hz : REAL;
    AccelRate_HzPerS : REAL := 20.0;
    DecelRate_HzPerS : REAL := 20.0; // Pente d'arret relevee sur trace reelle MES (-20.0 Hz/s)
    TimeConstant_S : REAL := 0.03;   // Reponse dynamique AC600 en boucle fermee (30 ms)
    LoadAngularVelocity_RadPerS : REAL;
    LoadFrequencyDroopGain_Hz : REAL := 0.50;
    CycleTime_S : REAL := 0.01;
END_VAR
VAR_OUTPUT
    Ready : BOOL;
    FrequencyCmd_Hz : REAL;
    ElectricalFrequency_Hz : REAL;
    ActualFrequency_Hz : REAL;
    ResponseAlpha : REAL;
END_VAR
VAR
    FrequencyDelta_Hz : REAL;
    FrequencyStep_Hz : REAL;
END_VAR
VAR CONSTANT
    CST_MinTime_S : REAL := 0.001;
    CST_StopFrequency_Hz : REAL := 0.5; // seuil nominal de fin de rampe variateur
    CST_MaxFrequency_Hz : REAL := 50.0; // plafond variateur reel (GVL_PERSISTENT._TranslationMaxFreq_Hz)
END_VAR

IF NOT Enable THEN
    Ready := FALSE;
    FrequencyCmd_Hz := 0.0;
    ElectricalFrequency_Hz := 0.0;
    ActualFrequency_Hz := 0.0;
    ResponseAlpha := 0.0;
    RETURN;
END_IF;

FrequencyDelta_Hz := LIMIT(0.0, FrequencyTgt_Hz, CST_MaxFrequency_Hz) - FrequencyCmd_Hz;
IF FrequencyDelta_Hz >= 0.0 THEN
    FrequencyStep_Hz := MAX(0.0, AccelRate_HzPerS) * CycleTime_S;
ELSE
    FrequencyStep_Hz := MAX(0.0, DecelRate_HzPerS) * CycleTime_S;
END_IF;
FrequencyCmd_Hz := FrequencyCmd_Hz + LIMIT(-FrequencyStep_Hz, FrequencyDelta_Hz, FrequencyStep_Hz);
IF TimeConstant_S > CST_MinTime_S THEN
    ResponseAlpha := CycleTime_S / (TimeConstant_S + CycleTime_S);
ELSE
    ResponseAlpha := 1.0;
END_IF;
ElectricalFrequency_Hz := ElectricalFrequency_Hz
    + ResponseAlpha * (FrequencyCmd_Hz - ElectricalFrequency_Hz);
(* Retour AC600 : frequence electrique de sortie. La charge est appliquee par le
   modele mecanique ; elle ne doit pas biaiser le retour publie au PLC. *)
ActualFrequency_Hz := MAX(0.0, ElectricalFrequency_Hz);
IF (FrequencyTgt_Hz <= 0.0) AND (FrequencyCmd_Hz <= 0.0)
    AND (ActualFrequency_Hz <= CST_StopFrequency_Hz) THEN
    ElectricalFrequency_Hz := 0.0;
    ActualFrequency_Hz := 0.0;
END_IF;
Ready := TRUE;
